(* IEC 61131-3 sources: REFUSR/GP/Refusr.jl/samples (part 13) *)

(* ---- 5-MUX_dozen-armor-usurp.st ---- *)
(*
This code implements a shuffled multiplexer with 5 control bits.
The control bits are: Data[N2], Data[N21], Data[N22], Data[N3], Data[N20]
The input bits are: Data[N24], Data[N4], Data[N27], Data[N1], Data[N23], Data[N25], Data[N5], Data[N26], Data[N31], Data[N7], Data[N8], Data[N6], Data[N9], Data[N28], Data[N13], Data[N11], Data[N12], Data[N29], Data[N30], Data[N33], Data[N10], Data[N34], Data[N35], Data[N37], Data[N32], Data[N14], Data[N16], Data[N36], Data[N17], Data[N18], Data[N19], Data[N15]

The symbolic expression is:
((((((((((((((((((((((((((((((((!(((((!(IN2)) & (!(IN21))) & (!(IN22))) & (!(IN3))) & (!(IN20)))) | IN24) & ((!((((IN2 & (!(IN21))) & (!(IN22))) & (!(IN3))) & (!(IN20)))) | IN4)) & ((!(((((!(IN2)) & IN21) & (!(IN22))) & (!(IN3))) & (!(IN20)))) | IN27)) & ((!((((IN2 & IN21) & (!(IN22))) & (!(IN3))) & (!(IN20)))) | IN1)) & ((!(((((!(IN2)) & (!(IN21))) & IN22) & (!(IN3))) & (!(IN20)))) | IN23)) & ((!((((IN2 & (!(IN21))) & IN22) & (!(IN3))) & (!(IN20)))) | IN25)) & ((!(((((!(IN2)) & IN21) & IN22) & (!(IN3))) & (!(IN20)))) | IN5)) & ((!((((IN2 & IN21) & IN22) & (!(IN3))) & (!(IN20)))) | IN26)) & ((!(((((!(IN2)) & (!(IN21))) & (!(IN22))) & IN3) & (!(IN20)))) | IN31)) & ((!((((IN2 & (!(IN21))) & (!(IN22))) & IN3) & (!(IN20)))) | IN7)) & ((!(((((!(IN2)) & IN21) & (!(IN22))) & IN3) & (!(IN20)))) | IN8)) & ((!((((IN2 & IN21) & (!(IN22))) & IN3) & (!(IN20)))) | IN6)) & ((!(((((!(IN2)) & (!(IN21))) & IN22) & IN3) & (!(IN20)))) | IN9)) & ((!((((IN2 & (!(IN21))) & IN22) & IN3) & (!(IN20)))) | IN28)) & ((!(((((!(IN2)) & IN21) & IN22) & IN3) & (!(IN20)))) | IN13)) & ((!((((IN2 & IN21) & IN22) & IN3) & (!(IN20)))) | IN11)) & ((!(((((!(IN2)) & (!(IN21))) & (!(IN22))) & (!(IN3))) & IN20)) | IN12)) & ((!((((IN2 & (!(IN21))) & (!(IN22))) & (!(IN3))) & IN20)) | IN29)) & ((!(((((!(IN2)) & IN21) & (!(IN22))) & (!(IN3))) & IN20)) | IN30)) & ((!((((IN2 & IN21) & (!(IN22))) & (!(IN3))) & IN20)) | IN33)) & ((!(((((!(IN2)) & (!(IN21))) & IN22) & (!(IN3))) & IN20)) | IN10)) & ((!((((IN2 & (!(IN21))) & IN22) & (!(IN3))) & IN20)) | IN34)) & ((!(((((!(IN2)) & IN21) & IN22) & (!(IN3))) & IN20)) | IN35)) & ((!((((IN2 & IN21) & IN22) & (!(IN3))) & IN20)) | IN37)) & ((!(((((!(IN2)) & (!(IN21))) & (!(IN22))) & IN3) & IN20)) | IN32)) & ((!((((IN2 & (!(IN21))) & (!(IN22))) & IN3) & IN20)) | IN14)) & ((!(((((!(IN2)) & IN21) & (!(IN22))) & IN3) & IN20)) | IN16)) & ((!((((IN2 & IN21) & (!(IN22))) & IN3) & IN20)) | IN36)) & ((!(((((!(IN2)) & (!(IN21))) & IN22) & IN3) & IN20)) | IN17)) & ((!((((IN2 & (!(IN21))) & IN22) & IN3) & IN20)) | IN18)) & ((!(((((!(IN2)) & IN21) & IN22) & IN3) & IN20)) | IN19)) & ((!((((IN2 & IN21) & IN22) & IN3) & IN20)) | IN15)

*)

FUNCTION_BLOCK F_CollectInput
  VAR_IN_OUT
      Data : ARRAY[1..40] OF BOOL;
  END_VAR
  VAR_INPUT
      TICK  : BOOL := 0;
      IN1   : BOOL := 0;
      IN2   : BOOL := 0;
      IN3   : BOOL := 0;
      IN4   : BOOL := 0;
      IN5   : BOOL := 0;
      RESET : BOOL := FALSE;
  END_VAR
  VAR_OUTPUT
      Finished : BOOL;
  END_VAR
  VAR
      j    : USINT := 1;
      tock : BOOL  := 0;
  END_VAR
  IF NOT RESET AND tock = NOT TICK THEN
      Data[j]   := IN1;
      Data[j+1] := IN2;
      Data[j+2] := IN3;
      Data[j+3] := IN4;
      Data[j+4] := IN5;
      j := j + 5;
      tock := TICK;
  ELSE
      j := 1;
      tock := 0;
  END_IF;
  Finished := (j > 40);
END_FUNCTION_BLOCK

PROGRAM Boiler
  VAR
    Data  : ARRAY[1..40] OF BOOL;
    Ready : BOOL;
    CollectInput : F_CollectInput;
  END_VAR
  VAR
    TICK     AT %IX1.0 : BOOL;
    IN1      AT %IX0.3 : BOOL;
    IN2      AT %IX0.4 : BOOL;
    IN3      AT %IX0.5 : BOOL;
    IN4      AT %IX0.6 : BOOL;
    IN5      AT %IX0.7 : BOOL;
    OutReady AT %QX0.0 : BOOL := FALSE;
    FeedNext AT %QX0.1 : BOOL := FALSE;
    Out      AT %QX0.2 : BOOL;
  END_VAR
  CollectInput(TICK:=TICK, IN1:=IN1, IN2:=IN2, IN3:=IN3, IN4:=IN4, IN5:=IN5);
  Ready := CollectInput.Finished;
  FeedNext := 1;
  IF Ready THEN
    Out := (((((((((((((((((((((((((((((((((NOT (((((NOT Data[2]) AND (NOT Data[21])) AND (NOT Data[22])) AND (NOT Data[3])) AND (NOT Data[20]))) OR Data[24]) AND ((NOT ((((Data[2] AND (NOT Data[21])) AND (NOT Data[22])) AND (NOT Data[3])) AND (NOT Data[20]))) OR Data[4])) AND ((NOT (((((NOT Data[2]) AND Data[21]) AND (NOT Data[22])) AND (NOT Data[3])) AND (NOT Data[20]))) OR Data[27])) AND ((NOT ((((Data[2] AND Data[21]) AND (NOT Data[22])) AND (NOT Data[3])) AND (NOT Data[20]))) OR Data[1])) AND ((NOT (((((NOT Data[2]) AND (NOT Data[21])) AND Data[22]) AND (NOT Data[3])) AND (NOT Data[20]))) OR Data[23])) AND ((NOT ((((Data[2] AND (NOT Data[21])) AND Data[22]) AND (NOT Data[3])) AND (NOT Data[20]))) OR Data[25])) AND ((NOT (((((NOT Data[2]) AND Data[21]) AND Data[22]) AND (NOT Data[3])) AND (NOT Data[20]))) OR Data[5])) AND ((NOT ((((Data[2] AND Data[21]) AND Data[22]) AND (NOT Data[3])) AND (NOT Data[20]))) OR Data[26])) AND ((NOT (((((NOT Data[2]) AND (NOT Data[21])) AND (NOT Data[22])) AND Data[3]) AND (NOT Data[20]))) OR Data[31])) AND ((NOT ((((Data[2] AND (NOT Data[21])) AND (NOT Data[22])) AND Data[3]) AND (NOT Data[20]))) OR Data[7])) AND ((NOT (((((NOT Data[2]) AND Data[21]) AND (NOT Data[22])) AND Data[3]) AND (NOT Data[20]))) OR Data[8])) AND ((NOT ((((Data[2] AND Data[21]) AND (NOT Data[22])) AND Data[3]) AND (NOT Data[20]))) OR Data[6])) AND ((NOT (((((NOT Data[2]) AND (NOT Data[21])) AND Data[22]) AND Data[3]) AND (NOT Data[20]))) OR Data[9])) AND ((NOT ((((Data[2] AND (NOT Data[21])) AND Data[22]) AND Data[3]) AND (NOT Data[20]))) OR Data[28])) AND ((NOT (((((NOT Data[2]) AND Data[21]) AND Data[22]) AND Data[3]) AND (NOT Data[20]))) OR Data[13])) AND ((NOT ((((Data[2] AND Data[21]) AND Data[22]) AND Data[3]) AND (NOT Data[20]))) OR Data[11])) AND ((NOT (((((NOT Data[2]) AND (NOT Data[21])) AND (NOT Data[22])) AND (NOT Data[3])) AND Data[20])) OR Data[12])) AND ((NOT ((((Data[2] AND (NOT Data[21])) AND (NOT Data[22])) AND (NOT Data[3])) AND Data[20])) OR Data[29])) AND ((NOT (((((NOT Data[2]) AND Data[21]) AND (NOT Data[22])) AND (NOT Data[3])) AND Data[20])) OR Data[30])) AND ((NOT ((((Data[2] AND Data[21]) AND (NOT Data[22])) AND (NOT Data[3])) AND Data[20])) OR Data[33])) AND ((NOT (((((NOT Data[2]) AND (NOT Data[21])) AND Data[22]) AND (NOT Data[3])) AND Data[20])) OR Data[10])) AND ((NOT ((((Data[2] AND (NOT Data[21])) AND Data[22]) AND (NOT Data[3])) AND Data[20])) OR Data[34])) AND ((NOT (((((NOT Data[2]) AND Data[21]) AND Data[22]) AND (NOT Data[3])) AND Data[20])) OR Data[35])) AND ((NOT ((((Data[2] AND Data[21]) AND Data[22]) AND (NOT Data[3])) AND Data[20])) OR Data[37])) AND ((NOT (((((NOT Data[2]) AND (NOT Data[21])) AND (NOT Data[22])) AND Data[3]) AND Data[20])) OR Data[32])) AND ((NOT ((((Data[2] AND (NOT Data[21])) AND (NOT Data[22])) AND Data[3]) AND Data[20])) OR Data[14])) AND ((NOT (((((NOT Data[2]) AND Data[21]) AND (NOT Data[22])) AND Data[3]) AND Data[20])) OR Data[16])) AND ((NOT ((((Data[2] AND Data[21]) AND (NOT Data[22])) AND Data[3]) AND Data[20])) OR Data[36])) AND ((NOT (((((NOT Data[2]) AND (NOT Data[21])) AND Data[22]) AND Data[3]) AND Data[20])) OR Data[17])) AND ((NOT ((((Data[2] AND (NOT Data[21])) AND Data[22]) AND Data[3]) AND Data[20])) OR Data[18])) AND ((NOT (((((NOT Data[2]) AND Data[21]) AND Data[22]) AND Data[3]) AND Data[20])) OR Data[19])) AND ((NOT ((((Data[2] AND Data[21]) AND Data[22]) AND Data[3]) AND Data[20])) OR Data[15]));
    OutReady := 1;
    CollectInput(RESET:=TRUE);
  END_IF;
END_PROGRAM

CONFIGURATION Config0
  RESOURCE Res0 ON PLC
    TASK task0(INTERVAL := T#20ms,PRIORITY := 0);
    PROGRAM instance0 WITH task0 : Boiler;
  END_RESOURCE
END_CONFIGURATION

(* ---- 5-MUX_froth-crick-hertz.st ---- *)
(*
This code implements a shuffled multiplexer with 5 control bits.
The control bits are: Data[N3], Data[N1], Data[N5], Data[N21], Data[N6]
The input bits are: Data[N4], Data[N20], Data[N2], Data[N7], Data[N22], Data[N8], Data[N10], Data[N11], Data[N13], Data[N26], Data[N23], Data[N25], Data[N9], Data[N14], Data[N24], Data[N29], Data[N16], Data[N27], Data[N15], Data[N12], Data[N17], Data[N19], Data[N32], Data[N30], Data[N28], Data[N18], Data[N31], Data[N33], Data[N37], Data[N35], Data[N36], Data[N34]

The symbolic expression is:
((((((((((((((((((((((((((((((((!(((((!(IN3)) & (!(IN1))) & (!(IN5))) & (!(IN21))) & (!(IN6)))) | IN4) & ((!((((IN3 & (!(IN1))) & (!(IN5))) & (!(IN21))) & (!(IN6)))) | IN20)) & ((!(((((!(IN3)) & IN1) & (!(IN5))) & (!(IN21))) & (!(IN6)))) | IN2)) & ((!((((IN3 & IN1) & (!(IN5))) & (!(IN21))) & (!(IN6)))) | IN7)) & ((!(((((!(IN3)) & (!(IN1))) & IN5) & (!(IN21))) & (!(IN6)))) | IN22)) & ((!((((IN3 & (!(IN1))) & IN5) & (!(IN21))) & (!(IN6)))) | IN8)) & ((!(((((!(IN3)) & IN1) & IN5) & (!(IN21))) & (!(IN6)))) | IN10)) & ((!((((IN3 & IN1) & IN5) & (!(IN21))) & (!(IN6)))) | IN11)) & ((!(((((!(IN3)) & (!(IN1))) & (!(IN5))) & IN21) & (!(IN6)))) | IN13)) & ((!((((IN3 & (!(IN1))) & (!(IN5))) & IN21) & (!(IN6)))) | IN26)) & ((!(((((!(IN3)) & IN1) & (!(IN5))) & IN21) & (!(IN6)))) | IN23)) & ((!((((IN3 & IN1) & (!(IN5))) & IN21) & (!(IN6)))) | IN25)) & ((!(((((!(IN3)) & (!(IN1))) & IN5) & IN21) & (!(IN6)))) | IN9)) & ((!((((IN3 & (!(IN1))) & IN5) & IN21) & (!(IN6)))) | IN14)) & ((!(((((!(IN3)) & IN1) & IN5) & IN21) & (!(IN6)))) | IN24)) & ((!((((IN3 & IN1) & IN5) & IN21) & (!(IN6)))) | IN29)) & ((!(((((!(IN3)) & (!(IN1))) & (!(IN5))) & (!(IN21))) & IN6)) | IN16)) & ((!((((IN3 & (!(IN1))) & (!(IN5))) & (!(IN21))) & IN6)) | IN27)) & ((!(((((!(IN3)) & IN1) & (!(IN5))) & (!(IN21))) & IN6)) | IN15)) & ((!((((IN3 & IN1) & (!(IN5))) & (!(IN21))) & IN6)) | IN12)) & ((!(((((!(IN3)) & (!(IN1))) & IN5) & (!(IN21))) & IN6)) | IN17)) & ((!((((IN3 & (!(IN1))) & IN5) & (!(IN21))) & IN6)) | IN19)) & ((!(((((!(IN3)) & IN1) & IN5) & (!(IN21))) & IN6)) | IN32)) & ((!((((IN3 & IN1) & IN5) & (!(IN21))) & IN6)) | IN30)) & ((!(((((!(IN3)) & (!(IN1))) & (!(IN5))) & IN21) & IN6)) | IN28)) & ((!((((IN3 & (!(IN1))) & (!(IN5))) & IN21) & IN6)) | IN18)) & ((!(((((!(IN3)) & IN1) & (!(IN5))) & IN21) & IN6)) | IN31)) & ((!((((IN3 & IN1) & (!(IN5))) & IN21) & IN6)) | IN33)) & ((!(((((!(IN3)) & (!(IN1))) & IN5) & IN21) & IN6)) | IN37)) & ((!((((IN3 & (!(IN1))) & IN5) & IN21) & IN6)) | IN35)) & ((!(((((!(IN3)) & IN1) & IN5) & IN21) & IN6)) | IN36)) & ((!((((IN3 & IN1) & IN5) & IN21) & IN6)) | IN34)

*)

FUNCTION_BLOCK F_CollectInput
  VAR_IN_OUT
      Data : ARRAY[1..40] OF BOOL;
  END_VAR
  VAR_INPUT
      TICK  : BOOL := 0;
      IN1   : BOOL := 0;
      IN2   : BOOL := 0;
      IN3   : BOOL := 0;
      IN4   : BOOL := 0;
      IN5   : BOOL := 0;
      RESET : BOOL := FALSE;
  END_VAR
  VAR_OUTPUT
      Finished : BOOL;
  END_VAR
  VAR
      j    : USINT := 1;
      tock : BOOL  := 0;
  END_VAR
  IF NOT RESET AND tock = NOT TICK THEN
      Data[j]   := IN1;
      Data[j+1] := IN2;
      Data[j+2] := IN3;
      Data[j+3] := IN4;
      Data[j+4] := IN5;
      j := j + 5;
      tock := TICK;
  ELSE
      j := 1;
      tock := 0;
  END_IF;
  Finished := (j > 40);
END_FUNCTION_BLOCK

PROGRAM Boiler
  VAR
    Data  : ARRAY[1..40] OF BOOL;
    Ready : BOOL;
    CollectInput : F_CollectInput;
  END_VAR
  VAR
    TICK     AT %IX1.0 : BOOL;
    IN1      AT %IX0.3 : BOOL;
    IN2      AT %IX0.4 : BOOL;
    IN3      AT %IX0.5 : BOOL;
    IN4      AT %IX0.6 : BOOL;
    IN5      AT %IX0.7 : BOOL;
    OutReady AT %QX0.0 : BOOL := FALSE;
    FeedNext AT %QX0.1 : BOOL := FALSE;
    Out      AT %QX0.2 : BOOL;
  END_VAR
  CollectInput(TICK:=TICK, IN1:=IN1, IN2:=IN2, IN3:=IN3, IN4:=IN4, IN5:=IN5);
  Ready := CollectInput.Finished;
  FeedNext := 1;
  IF Ready THEN
    Out := (((((((((((((((((((((((((((((((((NOT (((((NOT Data[3]) AND (NOT Data[1])) AND (NOT Data[5])) AND (NOT Data[21])) AND (NOT Data[6]))) OR Data[4]) AND ((NOT ((((Data[3] AND (NOT Data[1])) AND (NOT Data[5])) AND (NOT Data[21])) AND (NOT Data[6]))) OR Data[20])) AND ((NOT (((((NOT Data[3]) AND Data[1]) AND (NOT Data[5])) AND (NOT Data[21])) AND (NOT Data[6]))) OR Data[2])) AND ((NOT ((((Data[3] AND Data[1]) AND (NOT Data[5])) AND (NOT Data[21])) AND (NOT Data[6]))) OR Data[7])) AND ((NOT (((((NOT Data[3]) AND (NOT Data[1])) AND Data[5]) AND (NOT Data[21])) AND (NOT Data[6]))) OR Data[22])) AND ((NOT ((((Data[3] AND (NOT Data[1])) AND Data[5]) AND (NOT Data[21])) AND (NOT Data[6]))) OR Data[8])) AND ((NOT (((((NOT Data[3]) AND Data[1]) AND Data[5]) AND (NOT Data[21])) AND (NOT Data[6]))) OR Data[10])) AND ((NOT ((((Data[3] AND Data[1]) AND Data[5]) AND (NOT Data[21])) AND (NOT Data[6]))) OR Data[11])) AND ((NOT (((((NOT Data[3]) AND (NOT Data[1])) AND (NOT Data[5])) AND Data[21]) AND (NOT Data[6]))) OR Data[13])) AND ((NOT ((((Data[3] AND (NOT Data[1])) AND (NOT Data[5])) AND Data[21]) AND (NOT Data[6]))) OR Data[26])) AND ((NOT (((((NOT Data[3]) AND Data[1]) AND (NOT Data[5])) AND Data[21]) AND (NOT Data[6]))) OR Data[23])) AND ((NOT ((((Data[3] AND Data[1]) AND (NOT Data[5])) AND Data[21]) AND (NOT Data[6]))) OR Data[25])) AND ((NOT (((((NOT Data[3]) AND (NOT Data[1])) AND Data[5]) AND Data[21]) AND (NOT Data[6]))) OR Data[9])) AND ((NOT ((((Data[3] AND (NOT Data[1])) AND Data[5]) AND Data[21]) AND (NOT Data[6]))) OR Data[14])) AND ((NOT (((((NOT Data[3]) AND Data[1]) AND Data[5]) AND Data[21]) AND (NOT Data[6]))) OR Data[24])) AND ((NOT ((((Data[3] AND Data[1]) AND Data[5]) AND Data[21]) AND (NOT Data[6]))) OR Data[29])) AND ((NOT (((((NOT Data[3]) AND (NOT Data[1])) AND (NOT Data[5])) AND (NOT Data[21])) AND Data[6])) OR Data[16])) AND ((NOT ((((Data[3] AND (NOT Data[1])) AND (NOT Data[5])) AND (NOT Data[21])) AND Data[6])) OR Data[27])) AND ((NOT (((((NOT Data[3]) AND Data[1]) AND (NOT Data[5])) AND (NOT Data[21])) AND Data[6])) OR Data[15])) AND ((NOT ((((Data[3] AND Data[1]) AND (NOT Data[5])) AND (NOT Data[21])) AND Data[6])) OR Data[12])) AND ((NOT (((((NOT Data[3]) AND (NOT Data[1])) AND Data[5]) AND (NOT Data[21])) AND Data[6])) OR Data[17])) AND ((NOT ((((Data[3] AND (NOT Data[1])) AND Data[5]) AND (NOT Data[21])) AND Data[6])) OR Data[19])) AND ((NOT (((((NOT Data[3]) AND Data[1]) AND Data[5]) AND (NOT Data[21])) AND Data[6])) OR Data[32])) AND ((NOT ((((Data[3] AND Data[1]) AND Data[5]) AND (NOT Data[21])) AND Data[6])) OR Data[30])) AND ((NOT (((((NOT Data[3]) AND (NOT Data[1])) AND (NOT Data[5])) AND Data[21]) AND Data[6])) OR Data[28])) AND ((NOT ((((Data[3] AND (NOT Data[1])) AND (NOT Data[5])) AND Data[21]) AND Data[6])) OR Data[18])) AND ((NOT (((((NOT Data[3]) AND Data[1]) AND (NOT Data[5])) AND Data[21]) AND Data[6])) OR Data[31])) AND ((NOT ((((Data[3] AND Data[1]) AND (NOT Data[5])) AND Data[21]) AND Data[6])) OR Data[33])) AND ((NOT (((((NOT Data[3]) AND (NOT Data[1])) AND Data[5]) AND Data[21]) AND Data[6])) OR Data[37])) AND ((NOT ((((Data[3] AND (NOT Data[1])) AND Data[5]) AND Data[21]) AND Data[6])) OR Data[35])) AND ((NOT (((((NOT Data[3]) AND Data[1]) AND Data[5]) AND Data[21]) AND Data[6])) OR Data[36])) AND ((NOT ((((Data[3] AND Data[1]) AND Data[5]) AND Data[21]) AND Data[6])) OR Data[34]));
    OutReady := 1;
    CollectInput(RESET:=TRUE);
  END_IF;
END_PROGRAM

CONFIGURATION Config0
  RESOURCE Res0 ON PLC
    TASK task0(INTERVAL := T#20ms,PRIORITY := 0);
    PROGRAM instance0 WITH task0 : Boiler;
  END_RESOURCE
END_CONFIGURATION

(* ---- 5-MUX_funds-axman-titan.st ---- *)
(*
This code implements a shuffled multiplexer with 5 control bits.
The control bits are: Data[N22], Data[N1], Data[N23], Data[N20], Data[N24]
The input bits are: Data[N26], Data[N21], Data[N29], Data[N27], Data[N7], Data[N4], Data[N30], Data[N33], Data[N25], Data[N28], Data[N31], Data[N34], Data[N6], Data[N2], Data[N32], Data[N8], Data[N3], Data[N14], Data[N9], Data[N5], Data[N10], Data[N35], Data[N12], Data[N13], Data[N16], Data[N15], Data[N36], Data[N37], Data[N11], Data[N17], Data[N19], Data[N18]

The symbolic expression is:
((((((((((((((((((((((((((((((((!(((((!(IN22)) & (!(IN1))) & (!(IN23))) & (!(IN20))) & (!(IN24)))) | IN26) & ((!((((IN22 & (!(IN1))) & (!(IN23))) & (!(IN20))) & (!(IN24)))) | IN21)) & ((!(((((!(IN22)) & IN1) & (!(IN23))) & (!(IN20))) & (!(IN24)))) | IN29)) & ((!((((IN22 & IN1) & (!(IN23))) & (!(IN20))) & (!(IN24)))) | IN27)) & ((!(((((!(IN22)) & (!(IN1))) & IN23) & (!(IN20))) & (!(IN24)))) | IN7)) & ((!((((IN22 & (!(IN1))) & IN23) & (!(IN20))) & (!(IN24)))) | IN4)) & ((!(((((!(IN22)) & IN1) & IN23) & (!(IN20))) & (!(IN24)))) | IN30)) & ((!((((IN22 & IN1) & IN23) & (!(IN20))) & (!(IN24)))) | IN33)) & ((!(((((!(IN22)) & (!(IN1))) & (!(IN23))) & IN20) & (!(IN24)))) | IN25)) & ((!((((IN22 & (!(IN1))) & (!(IN23))) & IN20) & (!(IN24)))) | IN28)) & ((!(((((!(IN22)) & IN1) & (!(IN23))) & IN20) & (!(IN24)))) | IN31)) & ((!((((IN22 & IN1) & (!(IN23))) & IN20) & (!(IN24)))) | IN34)) & ((!(((((!(IN22)) & (!(IN1))) & IN23) & IN20) & (!(IN24)))) | IN6)) & ((!((((IN22 & (!(IN1))) & IN23) & IN20) & (!(IN24)))) | IN2)) & ((!(((((!(IN22)) & IN1) & IN23) & IN20) & (!(IN24)))) | IN32)) & ((!((((IN22 & IN1) & IN23) & IN20) & (!(IN24)))) | IN8)) & ((!(((((!(IN22)) & (!(IN1))) & (!(IN23))) & (!(IN20))) & IN24)) | IN3)) & ((!((((IN22 & (!(IN1))) & (!(IN23))) & (!(IN20))) & IN24)) | IN14)) & ((!(((((!(IN22)) & IN1) & (!(IN23))) & (!(IN20))) & IN24)) | IN9)) & ((!((((IN22 & IN1) & (!(IN23))) & (!(IN20))) & IN24)) | IN5)) & ((!(((((!(IN22)) & (!(IN1))) & IN23) & (!(IN20))) & IN24)) | IN10)) & ((!((((IN22 & (!(IN1))) & IN23) & (!(IN20))) & IN24)) | IN35)) & ((!(((((!(IN22)) & IN1) & IN23) & (!(IN20))) & IN24)) | IN12)) & ((!((((IN22 & IN1) & IN23) & (!(IN20))) & IN24)) | IN13)) & ((!(((((!(IN22)) & (!(IN1))) & (!(IN23))) & IN20) & IN24)) | IN16)) & ((!((((IN22 & (!(IN1))) & (!(IN23))) & IN20) & IN24)) | IN15)) & ((!(((((!(IN22)) & IN1) & (!(IN23))) & IN20) & IN24)) | IN36)) & ((!((((IN22 & IN1) & (!(IN23))) & IN20) & IN24)) | IN37)) & ((!(((((!(IN22)) & (!(IN1))) & IN23) & IN20) & IN24)) | IN11)) & ((!((((IN22 & (!(IN1))) & IN23) & IN20) & IN24)) | IN17)) & ((!(((((!(IN22)) & IN1) & IN23) & IN20) & IN24)) | IN19)) & ((!((((IN22 & IN1) & IN23) & IN20) & IN24)) | IN18)

*)

FUNCTION_BLOCK F_CollectInput
  VAR_IN_OUT
      Data : ARRAY[1..40] OF BOOL;
  END_VAR
  VAR_INPUT
      TICK  : BOOL := 0;
      IN1   : BOOL := 0;
      IN2   : BOOL := 0;
      IN3   : BOOL := 0;
      IN4   : BOOL := 0;
      IN5   : BOOL := 0;
      RESET : BOOL := FALSE;
  END_VAR
  VAR_OUTPUT
      Finished : BOOL;
  END_VAR
  VAR
      j    : USINT := 1;
      tock : BOOL  := 0;
  END_VAR
  IF NOT RESET AND tock = NOT TICK THEN
      Data[j]   := IN1;
      Data[j+1] := IN2;
      Data[j+2] := IN3;
      Data[j+3] := IN4;
      Data[j+4] := IN5;
      j := j + 5;
      tock := TICK;
  ELSE
      j := 1;
      tock := 0;
  END_IF;
  Finished := (j > 40);
END_FUNCTION_BLOCK

PROGRAM Boiler
  VAR
    Data  : ARRAY[1..40] OF BOOL;
    Ready : BOOL;
    CollectInput : F_CollectInput;
  END_VAR
  VAR
    TICK     AT %IX1.0 : BOOL;
    IN1      AT %IX0.3 : BOOL;
    IN2      AT %IX0.4 : BOOL;
    IN3      AT %IX0.5 : BOOL;
    IN4      AT %IX0.6 : BOOL;
    IN5      AT %IX0.7 : BOOL;
    OutReady AT %QX0.0 : BOOL := FALSE;
    FeedNext AT %QX0.1 : BOOL := FALSE;
    Out      AT %QX0.2 : BOOL;
  END_VAR
  CollectInput(TICK:=TICK, IN1:=IN1, IN2:=IN2, IN3:=IN3, IN4:=IN4, IN5:=IN5);
  Ready := CollectInput.Finished;
  FeedNext := 1;
  IF Ready THEN
    Out := (((((((((((((((((((((((((((((((((NOT (((((NOT Data[22]) AND (NOT Data[1])) AND (NOT Data[23])) AND (NOT Data[20])) AND (NOT Data[24]))) OR Data[26]) AND ((NOT ((((Data[22] AND (NOT Data[1])) AND (NOT Data[23])) AND (NOT Data[20])) AND (NOT Data[24]))) OR Data[21])) AND ((NOT (((((NOT Data[22]) AND Data[1]) AND (NOT Data[23])) AND (NOT Data[20])) AND (NOT Data[24]))) OR Data[29])) AND ((NOT ((((Data[22] AND Data[1]) AND (NOT Data[23])) AND (NOT Data[20])) AND (NOT Data[24]))) OR Data[27])) AND ((NOT (((((NOT Data[22]) AND (NOT Data[1])) AND Data[23]) AND (NOT Data[20])) AND (NOT Data[24]))) OR Data[7])) AND ((NOT ((((Data[22] AND (NOT Data[1])) AND Data[23]) AND (NOT Data[20])) AND (NOT Data[24]))) OR Data[4])) AND ((NOT (((((NOT Data[22]) AND Data[1]) AND Data[23]) AND (NOT Data[20])) AND (NOT Data[24]))) OR Data[30])) AND ((NOT ((((Data[22] AND Data[1]) AND Data[23]) AND (NOT Data[20])) AND (NOT Data[24]))) OR Data[33])) AND ((NOT (((((NOT Data[22]) AND (NOT Data[1])) AND (NOT Data[23])) AND Data[20]) AND (NOT Data[24]))) OR Data[25])) AND ((NOT ((((Data[22] AND (NOT Data[1])) AND (NOT Data[23])) AND Data[20]) AND (NOT Data[24]))) OR Data[28])) AND ((NOT (((((NOT Data[22]) AND Data[1]) AND (NOT Data[23])) AND Data[20]) AND (NOT Data[24]))) OR Data[31])) AND ((NOT ((((Data[22] AND Data[1]) AND (NOT Data[23])) AND Data[20]) AND (NOT Data[24]))) OR Data[34])) AND ((NOT (((((NOT Data[22]) AND (NOT Data[1])) AND Data[23]) AND Data[20]) AND (NOT Data[24]))) OR Data[6])) AND ((NOT ((((Data[22] AND (NOT Data[1])) AND Data[23]) AND Data[20]) AND (NOT Data[24]))) OR Data[2])) AND ((NOT (((((NOT Data[22]) AND Data[1]) AND Data[23]) AND Data[20]) AND (NOT Data[24]))) OR Data[32])) AND ((NOT ((((Data[22] AND Data[1]) AND Data[23]) AND Data[20]) AND (NOT Data[24]))) OR Data[8])) AND ((NOT (((((NOT Data[22]) AND (NOT Data[1])) AND (NOT Data[23])) AND (NOT Data[20])) AND Data[24])) OR Data[3])) AND ((NOT ((((Data[22] AND (NOT Data[1])) AND (NOT Data[23])) AND (NOT Data[20])) AND Data[24])) OR Data[14])) AND ((NOT (((((NOT Data[22]) AND Data[1]) AND (NOT Data[23])) AND (NOT Data[20])) AND Data[24])) OR Data[9])) AND ((NOT ((((Data[22] AND Data[1]) AND (NOT Data[23])) AND (NOT Data[20])) AND Data[24])) OR Data[5])) AND ((NOT (((((NOT Data[22]) AND (NOT Data[1])) AND Data[23]) AND (NOT Data[20])) AND Data[24])) OR Data[10])) AND ((NOT ((((Data[22] AND (NOT Data[1])) AND Data[23]) AND (NOT Data[20])) AND Data[24])) OR Data[35])) AND ((NOT (((((NOT Data[22]) AND Data[1]) AND Data[23]) AND (NOT Data[20])) AND Data[24])) OR Data[12])) AND ((NOT ((((Data[22] AND Data[1]) AND Data[23]) AND (NOT Data[20])) AND Data[24])) OR Data[13])) AND ((NOT (((((NOT Data[22]) AND (NOT Data[1])) AND (NOT Data[23])) AND Data[20]) AND Data[24])) OR Data[16])) AND ((NOT ((((Data[22] AND (NOT Data[1])) AND (NOT Data[23])) AND Data[20]) AND Data[24])) OR Data[15])) AND ((NOT (((((NOT Data[22]) AND Data[1]) AND (NOT Data[23])) AND Data[20]) AND Data[24])) OR Data[36])) AND ((NOT ((((Data[22] AND Data[1]) AND (NOT Data[23])) AND Data[20]) AND Data[24])) OR Data[37])) AND ((NOT (((((NOT Data[22]) AND (NOT Data[1])) AND Data[23]) AND Data[20]) AND Data[24])) OR Data[11])) AND ((NOT ((((Data[22] AND (NOT Data[1])) AND Data[23]) AND Data[20]) AND Data[24])) OR Data[17])) AND ((NOT (((((NOT Data[22]) AND Data[1]) AND Data[23]) AND Data[20]) AND Data[24])) OR Data[19])) AND ((NOT ((((Data[22] AND Data[1]) AND Data[23]) AND Data[20]) AND Data[24])) OR Data[18]));
    OutReady := 1;
    CollectInput(RESET:=TRUE);
  END_IF;
END_PROGRAM

CONFIGURATION Config0
  RESOURCE Res0 ON PLC
    TASK task0(INTERVAL := T#20ms,PRIORITY := 0);
    PROGRAM instance0 WITH task0 : Boiler;
  END_RESOURCE
END_CONFIGURATION

(* ---- 5-MUX_fungi-exalt-steer.st ---- *)
(*
This code implements a shuffled multiplexer with 5 control bits.
The control bits are: Data[N1], Data[N3], Data[N5], Data[N2], Data[N21]
The input bits are: Data[N20], Data[N25], Data[N6], Data[N23], Data[N26], Data[N24], Data[N4], Data[N13], Data[N28], Data[N7], Data[N22], Data[N29], Data[N30], Data[N27], Data[N10], Data[N11], Data[N31], Data[N33], Data[N34], Data[N32], Data[N8], Data[N36], Data[N35], Data[N37], Data[N15], Data[N17], Data[N14], Data[N9], Data[N12], Data[N18], Data[N16], Data[N19]

The symbolic expression is:
((((((((((((((((((((((((((((((((!(((((!(IN1)) & (!(IN3))) & (!(IN5))) & (!(IN2))) & (!(IN21)))) | IN20) & ((!((((IN1 & (!(IN3))) & (!(IN5))) & (!(IN2))) & (!(IN21)))) | IN25)) & ((!(((((!(IN1)) & IN3) & (!(IN5))) & (!(IN2))) & (!(IN21)))) | IN6)) & ((!((((IN1 & IN3) & (!(IN5))) & (!(IN2))) & (!(IN21)))) | IN23)) & ((!(((((!(IN1)) & (!(IN3))) & IN5) & (!(IN2))) & (!(IN21)))) | IN26)) & ((!((((IN1 & (!(IN3))) & IN5) & (!(IN2))) & (!(IN21)))) | IN24)) & ((!(((((!(IN1)) & IN3) & IN5) & (!(IN2))) & (!(IN21)))) | IN4)) & ((!((((IN1 & IN3) & IN5) & (!(IN2))) & (!(IN21)))) | IN13)) & ((!(((((!(IN1)) & (!(IN3))) & (!(IN5))) & IN2) & (!(IN21)))) | IN28)) & ((!((((IN1 & (!(IN3))) & (!(IN5))) & IN2) & (!(IN21)))) | IN7)) & ((!(((((!(IN1)) & IN3) & (!(IN5))) & IN2) & (!(IN21)))) | IN22)) & ((!((((IN1 & IN3) & (!(IN5))) & IN2) & (!(IN21)))) | IN29)) & ((!(((((!(IN1)) & (!(IN3))) & IN5) & IN2) & (!(IN21)))) | IN30)) & ((!((((IN1 & (!(IN3))) & IN5) & IN2) & (!(IN21)))) | IN27)) & ((!(((((!(IN1)) & IN3) & IN5) & IN2) & (!(IN21)))) | IN10)) & ((!((((IN1 & IN3) & IN5) & IN2) & (!(IN21)))) | IN11)) & ((!(((((!(IN1)) & (!(IN3))) & (!(IN5))) & (!(IN2))) & IN21)) | IN31)) & ((!((((IN1 & (!(IN3))) & (!(IN5))) & (!(IN2))) & IN21)) | IN33)) & ((!(((((!(IN1)) & IN3) & (!(IN5))) & (!(IN2))) & IN21)) | IN34)) & ((!((((IN1 & IN3) & (!(IN5))) & (!(IN2))) & IN21)) | IN32)) & ((!(((((!(IN1)) & (!(IN3))) & IN5) & (!(IN2))) & IN21)) | IN8)) & ((!((((IN1 & (!(IN3))) & IN5) & (!(IN2))) & IN21)) | IN36)) & ((!(((((!(IN1)) & IN3) & IN5) & (!(IN2))) & IN21)) | IN35)) & ((!((((IN1 & IN3) & IN5) & (!(IN2))) & IN21)) | IN37)) & ((!(((((!(IN1)) & (!(IN3))) & (!(IN5))) & IN2) & IN21)) | IN15)) & ((!((((IN1 & (!(IN3))) & (!(IN5))) & IN2) & IN21)) | IN17)) & ((!(((((!(IN1)) & IN3) & (!(IN5))) & IN2) & IN21)) | IN14)) & ((!((((IN1 & IN3) & (!(IN5))) & IN2) & IN21)) | IN9)) & ((!(((((!(IN1)) & (!(IN3))) & IN5) & IN2) & IN21)) | IN12)) & ((!((((IN1 & (!(IN3))) & IN5) & IN2) & IN21)) | IN18)) & ((!(((((!(IN1)) & IN3) & IN5) & IN2) & IN21)) | IN16)) & ((!((((IN1 & IN3) & IN5) & IN2) & IN21)) | IN19)

*)

FUNCTION_BLOCK F_CollectInput
  VAR_IN_OUT
      Data : ARRAY[1..40] OF BOOL;
  END_VAR
  VAR_INPUT
      TICK  : BOOL := 0;
      IN1   : BOOL := 0;
      IN2   : BOOL := 0;
      IN3   : BOOL := 0;
      IN4   : BOOL := 0;
      IN5   : BOOL := 0;
      RESET : BOOL := FALSE;
  END_VAR
  VAR_OUTPUT
      Finished : BOOL;
  END_VAR
  VAR
      j    : USINT := 1;
      tock : BOOL  := 0;
  END_VAR
  IF NOT RESET AND tock = NOT TICK THEN
      Data[j]   := IN1;
      Data[j+1] := IN2;
      Data[j+2] := IN3;
      Data[j+3] := IN4;
      Data[j+4] := IN5;
      j := j + 5;
      tock := TICK;
  ELSE
      j := 1;
      tock := 0;
  END_IF;
  Finished := (j > 40);
END_FUNCTION_BLOCK

PROGRAM Boiler
  VAR
    Data  : ARRAY[1..40] OF BOOL;
    Ready : BOOL;
    CollectInput : F_CollectInput;
  END_VAR
  VAR
    TICK     AT %IX1.0 : BOOL;
    IN1      AT %IX0.3 : BOOL;
    IN2      AT %IX0.4 : BOOL;
    IN3      AT %IX0.5 : BOOL;
    IN4      AT %IX0.6 : BOOL;
    IN5      AT %IX0.7 : BOOL;
    OutReady AT %QX0.0 : BOOL := FALSE;
    FeedNext AT %QX0.1 : BOOL := FALSE;
    Out      AT %QX0.2 : BOOL;
  END_VAR
  CollectInput(TICK:=TICK, IN1:=IN1, IN2:=IN2, IN3:=IN3, IN4:=IN4, IN5:=IN5);
  Ready := CollectInput.Finished;
  FeedNext := 1;
  IF Ready THEN
    Out := (((((((((((((((((((((((((((((((((NOT (((((NOT Data[1]) AND (NOT Data[3])) AND (NOT Data[5])) AND (NOT Data[2])) AND (NOT Data[21]))) OR Data[20]) AND ((NOT ((((Data[1] AND (NOT Data[3])) AND (NOT Data[5])) AND (NOT Data[2])) AND (NOT Data[21]))) OR Data[25])) AND ((NOT (((((NOT Data[1]) AND Data[3]) AND (NOT Data[5])) AND (NOT Data[2])) AND (NOT Data[21]))) OR Data[6])) AND ((NOT ((((Data[1] AND Data[3]) AND (NOT Data[5])) AND (NOT Data[2])) AND (NOT Data[21]))) OR Data[23])) AND ((NOT (((((NOT Data[1]) AND (NOT Data[3])) AND Data[5]) AND (NOT Data[2])) AND (NOT Data[21]))) OR Data[26])) AND ((NOT ((((Data[1] AND (NOT Data[3])) AND Data[5]) AND (NOT Data[2])) AND (NOT Data[21]))) OR Data[24])) AND ((NOT (((((NOT Data[1]) AND Data[3]) AND Data[5]) AND (NOT Data[2])) AND (NOT Data[21]))) OR Data[4])) AND ((NOT ((((Data[1] AND Data[3]) AND Data[5]) AND (NOT Data[2])) AND (NOT Data[21]))) OR Data[13])) AND ((NOT (((((NOT Data[1]) AND (NOT Data[3])) AND (NOT Data[5])) AND Data[2]) AND (NOT Data[21]))) OR Data[28])) AND ((NOT ((((Data[1] AND (NOT Data[3])) AND (NOT Data[5])) AND Data[2]) AND (NOT Data[21]))) OR Data[7])) AND ((NOT (((((NOT Data[1]) AND Data[3]) AND (NOT Data[5])) AND Data[2]) AND (NOT Data[21]))) OR Data[22])) AND ((NOT ((((Data[1] AND Data[3]) AND (NOT Data[5])) AND Data[2]) AND (NOT Data[21]))) OR Data[29])) AND ((NOT (((((NOT Data[1]) AND (NOT Data[3])) AND Data[5]) AND Data[2]) AND (NOT Data[21]))) OR Data[30])) AND ((NOT ((((Data[1] AND (NOT Data[3])) AND Data[5]) AND Data[2]) AND (NOT Data[21]))) OR Data[27])) AND ((NOT (((((NOT Data[1]) AND Data[3]) AND Data[5]) AND Data[2]) AND (NOT Data[21]))) OR Data[10])) AND ((NOT ((((Data[1] AND Data[3]) AND Data[5]) AND Data[2]) AND (NOT Data[21]))) OR Data[11])) AND ((NOT (((((NOT Data[1]) AND (NOT Data[3])) AND (NOT Data[5])) AND (NOT Data[2])) AND Data[21])) OR Data[31])) AND ((NOT ((((Data[1] AND (NOT Data[3])) AND (NOT Data[5])) AND (NOT Data[2])) AND Data[21])) OR Data[33])) AND ((NOT (((((NOT Data[1]) AND Data[3]) AND (NOT Data[5])) AND (NOT Data[2])) AND Data[21])) OR Data[34])) AND ((NOT ((((Data[1] AND Data[3]) AND (NOT Data[5])) AND (NOT Data[2])) AND Data[21])) OR Data[32])) AND ((NOT (((((NOT Data[1]) AND (NOT Data[3])) AND Data[5]) AND (NOT Data[2])) AND Data[21])) OR Data[8])) AND ((NOT ((((Data[1] AND (NOT Data[3])) AND Data[5]) AND (NOT Data[2])) AND Data[21])) OR Data[36])) AND ((NOT (((((NOT Data[1]) AND Data[3]) AND Data[5]) AND (NOT Data[2])) AND Data[21])) OR Data[35])) AND ((NOT ((((Data[1] AND Data[3]) AND Data[5]) AND (NOT Data[2])) AND Data[21])) OR Data[37])) AND ((NOT (((((NOT Data[1]) AND (NOT Data[3])) AND (NOT Data[5])) AND Data[2]) AND Data[21])) OR Data[15])) AND ((NOT ((((Data[1] AND (NOT Data[3])) AND (NOT Data[5])) AND Data[2]) AND Data[21])) OR Data[17])) AND ((NOT (((((NOT Data[1]) AND Data[3]) AND (NOT Data[5])) AND Data[2]) AND Data[21])) OR Data[14])) AND ((NOT ((((Data[1] AND Data[3]) AND (NOT Data[5])) AND Data[2]) AND Data[21])) OR Data[9])) AND ((NOT (((((NOT Data[1]) AND (NOT Data[3])) AND Data[5]) AND Data[2]) AND Data[21])) OR Data[12])) AND ((NOT ((((Data[1] AND (NOT Data[3])) AND Data[5]) AND Data[2]) AND Data[21])) OR Data[18])) AND ((NOT (((((NOT Data[1]) AND Data[3]) AND Data[5]) AND Data[2]) AND Data[21])) OR Data[16])) AND ((NOT ((((Data[1] AND Data[3]) AND Data[5]) AND Data[2]) AND Data[21])) OR Data[19]));
    OutReady := 1;
    CollectInput(RESET:=TRUE);
  END_IF;
END_PROGRAM

CONFIGURATION Config0
  RESOURCE Res0 ON PLC
    TASK task0(INTERVAL := T#20ms,PRIORITY := 0);
    PROGRAM instance0 WITH task0 : Boiler;
  END_RESOURCE
END_CONFIGURATION

(* ---- 5-MUX_gipsy-agave-shock.st ---- *)
(*
This code implements a shuffled multiplexer with 5 control bits.
The control bits are: Data[N21], Data[N23], Data[N24], Data[N25], Data[N26]
The input bits are: Data[N4], Data[N5], Data[N1], Data[N6], Data[N27], Data[N20], Data[N30], Data[N31], Data[N22], Data[N33], Data[N9], Data[N32], Data[N28], Data[N34], Data[N37], Data[N2], Data[N29], Data[N36], Data[N3], Data[N7], Data[N35], Data[N8], Data[N13], Data[N12], Data[N11], Data[N19], Data[N18], Data[N15], Data[N10], Data[N14], Data[N16], Data[N17]

The symbolic expression is:
((((((((((((((((((((((((((((((((!(((((!(IN21)) & (!(IN23))) & (!(IN24))) & (!(IN25))) & (!(IN26)))) | IN4) & ((!((((IN21 & (!(IN23))) & (!(IN24))) & (!(IN25))) & (!(IN26)))) | IN5)) & ((!(((((!(IN21)) & IN23) & (!(IN24))) & (!(IN25))) & (!(IN26)))) | IN1)) & ((!((((IN21 & IN23) & (!(IN24))) & (!(IN25))) & (!(IN26)))) | IN6)) & ((!(((((!(IN21)) & (!(IN23))) & IN24) & (!(IN25))) & (!(IN26)))) | IN27)) & ((!((((IN21 & (!(IN23))) & IN24) & (!(IN25))) & (!(IN26)))) | IN20)) & ((!(((((!(IN21)) & IN23) & IN24) & (!(IN25))) & (!(IN26)))) | IN30)) & ((!((((IN21 & IN23) & IN24) & (!(IN25))) & (!(IN26)))) | IN31)) & ((!(((((!(IN21)) & (!(IN23))) & (!(IN24))) & IN25) & (!(IN26)))) | IN22)) & ((!((((IN21 & (!(IN23))) & (!(IN24))) & IN25) & (!(IN26)))) | IN33)) & ((!(((((!(IN21)) & IN23) & (!(IN24))) & IN25) & (!(IN26)))) | IN9)) & ((!((((IN21 & IN23) & (!(IN24))) & IN25) & (!(IN26)))) | IN32)) & ((!(((((!(IN21)) & (!(IN23))) & IN24) & IN25) & (!(IN26)))) | IN28)) & ((!((((IN21 & (!(IN23))) & IN24) & IN25) & (!(IN26)))) | IN34)) & ((!(((((!(IN21)) & IN23) & IN24) & IN25) & (!(IN26)))) | IN37)) & ((!((((IN21 & IN23) & IN24) & IN25) & (!(IN26)))) | IN2)) & ((!(((((!(IN21)) & (!(IN23))) & (!(IN24))) & (!(IN25))) & IN26)) | IN29)) & ((!((((IN21 & (!(IN23))) & (!(IN24))) & (!(IN25))) & IN26)) | IN36)) & ((!(((((!(IN21)) & IN23) & (!(IN24))) & (!(IN25))) & IN26)) | IN3)) & ((!((((IN21 & IN23) & (!(IN24))) & (!(IN25))) & IN26)) | IN7)) & ((!(((((!(IN21)) & (!(IN23))) & IN24) & (!(IN25))) & IN26)) | IN35)) & ((!((((IN21 & (!(IN23))) & IN24) & (!(IN25))) & IN26)) | IN8)) & ((!(((((!(IN21)) & IN23) & IN24) & (!(IN25))) & IN26)) | IN13)) & ((!((((IN21 & IN23) & IN24) & (!(IN25))) & IN26)) | IN12)) & ((!(((((!(IN21)) & (!(IN23))) & (!(IN24))) & IN25) & IN26)) | IN11)) & ((!((((IN21 & (!(IN23))) & (!(IN24))) & IN25) & IN26)) | IN19)) & ((!(((((!(IN21)) & IN23) & (!(IN24))) & IN25) & IN26)) | IN18)) & ((!((((IN21 & IN23) & (!(IN24))) & IN25) & IN26)) | IN15)) & ((!(((((!(IN21)) & (!(IN23))) & IN24) & IN25) & IN26)) | IN10)) & ((!((((IN21 & (!(IN23))) & IN24) & IN25) & IN26)) | IN14)) & ((!(((((!(IN21)) & IN23) & IN24) & IN25) & IN26)) | IN16)) & ((!((((IN21 & IN23) & IN24) & IN25) & IN26)) | IN17)

*)

FUNCTION_BLOCK F_CollectInput
  VAR_IN_OUT
      Data : ARRAY[1..40] OF BOOL;
  END_VAR
  VAR_INPUT
      TICK  : BOOL := 0;
      IN1   : BOOL := 0;
      IN2   : BOOL := 0;
      IN3   : BOOL := 0;
      IN4   : BOOL := 0;
      IN5   : BOOL := 0;
      RESET : BOOL := FALSE;
  END_VAR
  VAR_OUTPUT
      Finished : BOOL;
  END_VAR
  VAR
      j    : USINT := 1;
      tock : BOOL  := 0;
  END_VAR
  IF NOT RESET AND tock = NOT TICK THEN
      Data[j]   := IN1;
      Data[j+1] := IN2;
      Data[j+2] := IN3;
      Data[j+3] := IN4;
      Data[j+4] := IN5;
      j := j + 5;
      tock := TICK;
  ELSE
      j := 1;
      tock := 0;
  END_IF;
  Finished := (j > 40);
END_FUNCTION_BLOCK

PROGRAM Boiler
  VAR
    Data  : ARRAY[1..40] OF BOOL;
    Ready : BOOL;
    CollectInput : F_CollectInput;
  END_VAR
  VAR
    TICK     AT %IX1.0 : BOOL;
    IN1      AT %IX0.3 : BOOL;
    IN2      AT %IX0.4 : BOOL;
    IN3      AT %IX0.5 : BOOL;
    IN4      AT %IX0.6 : BOOL;
    IN5      AT %IX0.7 : BOOL;
    OutReady AT %QX0.0 : BOOL := FALSE;
    FeedNext AT %QX0.1 : BOOL := FALSE;
    Out      AT %QX0.2 : BOOL;
  END_VAR
  CollectInput(TICK:=TICK, IN1:=IN1, IN2:=IN2, IN3:=IN3, IN4:=IN4, IN5:=IN5);
  Ready := CollectInput.Finished;
  FeedNext := 1;
  IF Ready THEN
    Out := (((((((((((((((((((((((((((((((((NOT (((((NOT Data[21]) AND (NOT Data[23])) AND (NOT Data[24])) AND (NOT Data[25])) AND (NOT Data[26]))) OR Data[4]) AND ((NOT ((((Data[21] AND (NOT Data[23])) AND (NOT Data[24])) AND (NOT Data[25])) AND (NOT Data[26]))) OR Data[5])) AND ((NOT (((((NOT Data[21]) AND Data[23]) AND (NOT Data[24])) AND (NOT Data[25])) AND (NOT Data[26]))) OR Data[1])) AND ((NOT ((((Data[21] AND Data[23]) AND (NOT Data[24])) AND (NOT Data[25])) AND (NOT Data[26]))) OR Data[6])) AND ((NOT (((((NOT Data[21]) AND (NOT Data[23])) AND Data[24]) AND (NOT Data[25])) AND (NOT Data[26]))) OR Data[27])) AND ((NOT ((((Data[21] AND (NOT Data[23])) AND Data[24]) AND (NOT Data[25])) AND (NOT Data[26]))) OR Data[20])) AND ((NOT (((((NOT Data[21]) AND Data[23]) AND Data[24]) AND (NOT Data[25])) AND (NOT Data[26]))) OR Data[30])) AND ((NOT ((((Data[21] AND Data[23]) AND Data[24]) AND (NOT Data[25])) AND (NOT Data[26]))) OR Data[31])) AND ((NOT (((((NOT Data[21]) AND (NOT Data[23])) AND (NOT Data[24])) AND Data[25]) AND (NOT Data[26]))) OR Data[22])) AND ((NOT ((((Data[21] AND (NOT Data[23])) AND (NOT Data[24])) AND Data[25]) AND (NOT Data[26]))) OR Data[33])) AND ((NOT (((((NOT Data[21]) AND Data[23]) AND (NOT Data[24])) AND Data[25]) AND (NOT Data[26]))) OR Data[9])) AND ((NOT ((((Data[21] AND Data[23]) AND (NOT Data[24])) AND Data[25]) AND (NOT Data[26]))) OR Data[32])) AND ((NOT (((((NOT Data[21]) AND (NOT Data[23])) AND Data[24]) AND Data[25]) AND (NOT Data[26]))) OR Data[28])) AND ((NOT ((((Data[21] AND (NOT Data[23])) AND Data[24]) AND Data[25]) AND (NOT Data[26]))) OR Data[34])) AND ((NOT (((((NOT Data[21]) AND Data[23]) AND Data[24]) AND Data[25]) AND (NOT Data[26]))) OR Data[37])) AND ((NOT ((((Data[21] AND Data[23]) AND Data[24]) AND Data[25]) AND (NOT Data[26]))) OR Data[2])) AND ((NOT (((((NOT Data[21]) AND (NOT Data[23])) AND (NOT Data[24])) AND (NOT Data[25])) AND Data[26])) OR Data[29])) AND ((NOT ((((Data[21] AND (NOT Data[23])) AND (NOT Data[24])) AND (NOT Data[25])) AND Data[26])) OR Data[36])) AND ((NOT (((((NOT Data[21]) AND Data[23]) AND (NOT Data[24])) AND (NOT Data[25])) AND Data[26])) OR Data[3])) AND ((NOT ((((Data[21] AND Data[23]) AND (NOT Data[24])) AND (NOT Data[25])) AND Data[26])) OR Data[7])) AND ((NOT (((((NOT Data[21]) AND (NOT Data[23])) AND Data[24]) AND (NOT Data[25])) AND Data[26])) OR Data[35])) AND ((NOT ((((Data[21] AND (NOT Data[23])) AND Data[24]) AND (NOT Data[25])) AND Data[26])) OR Data[8])) AND ((NOT (((((NOT Data[21]) AND Data[23]) AND Data[24]) AND (NOT Data[25])) AND Data[26])) OR Data[13])) AND ((NOT ((((Data[21] AND Data[23]) AND Data[24]) AND (NOT Data[25])) AND Data[26])) OR Data[12])) AND ((NOT (((((NOT Data[21]) AND (NOT Data[23])) AND (NOT Data[24])) AND Data[25]) AND Data[26])) OR Data[11])) AND ((NOT ((((Data[21] AND (NOT Data[23])) AND (NOT Data[24])) AND Data[25]) AND Data[26])) OR Data[19])) AND ((NOT (((((NOT Data[21]) AND Data[23]) AND (NOT Data[24])) AND Data[25]) AND Data[26])) OR Data[18])) AND ((NOT ((((Data[21] AND Data[23]) AND (NOT Data[24])) AND Data[25]) AND Data[26])) OR Data[15])) AND ((NOT (((((NOT Data[21]) AND (NOT Data[23])) AND Data[24]) AND Data[25]) AND Data[26])) OR Data[10])) AND ((NOT ((((Data[21] AND (NOT Data[23])) AND Data[24]) AND Data[25]) AND Data[26])) OR Data[14])) AND ((NOT (((((NOT Data[21]) AND Data[23]) AND Data[24]) AND Data[25]) AND Data[26])) OR Data[16])) AND ((NOT ((((Data[21] AND Data[23]) AND Data[24]) AND Data[25]) AND Data[26])) OR Data[17]));
    OutReady := 1;
    CollectInput(RESET:=TRUE);
  END_IF;
END_PROGRAM

CONFIGURATION Config0
  RESOURCE Res0 ON PLC
    TASK task0(INTERVAL := T#20ms,PRIORITY := 0);
    PROGRAM instance0 WITH task0 : Boiler;
  END_RESOURCE
END_CONFIGURATION

(* ---- 5-MUX_gloms-friar-gimme.st ---- *)
(*
This code implements a shuffled multiplexer with 5 control bits.
The control bits are: Data[N23], Data[N2], Data[N20], Data[N3], Data[N4]
The input bits are: Data[N21], Data[N26], Data[N1], Data[N22], Data[N25], Data[N24], Data[N5], Data[N6], Data[N31], Data[N33], Data[N8], Data[N27], Data[N30], Data[N29], Data[N9], Data[N32], Data[N12], Data[N10], Data[N28], Data[N7], Data[N13], Data[N14], Data[N11], Data[N34], Data[N35], Data[N37], Data[N15], Data[N16], Data[N36], Data[N17], Data[N18], Data[N19]

The symbolic expression is:
((((((((((((((((((((((((((((((((!(((((!(IN23)) & (!(IN2))) & (!(IN20))) & (!(IN3))) & (!(IN4)))) | IN21) & ((!((((IN23 & (!(IN2))) & (!(IN20))) & (!(IN3))) & (!(IN4)))) | IN26)) & ((!(((((!(IN23)) & IN2) & (!(IN20))) & (!(IN3))) & (!(IN4)))) | IN1)) & ((!((((IN23 & IN2) & (!(IN20))) & (!(IN3))) & (!(IN4)))) | IN22)) & ((!(((((!(IN23)) & (!(IN2))) & IN20) & (!(IN3))) & (!(IN4)))) | IN25)) & ((!((((IN23 & (!(IN2))) & IN20) & (!(IN3))) & (!(IN4)))) | IN24)) & ((!(((((!(IN23)) & IN2) & IN20) & (!(IN3))) & (!(IN4)))) | IN5)) & ((!((((IN23 & IN2) & IN20) & (!(IN3))) & (!(IN4)))) | IN6)) & ((!(((((!(IN23)) & (!(IN2))) & (!(IN20))) & IN3) & (!(IN4)))) | IN31)) & ((!((((IN23 & (!(IN2))) & (!(IN20))) & IN3) & (!(IN4)))) | IN33)) & ((!(((((!(IN23)) & IN2) & (!(IN20))) & IN3) & (!(IN4)))) | IN8)) & ((!((((IN23 & IN2) & (!(IN20))) & IN3) & (!(IN4)))) | IN27)) & ((!(((((!(IN23)) & (!(IN2))) & IN20) & IN3) & (!(IN4)))) | IN30)) & ((!((((IN23 & (!(IN2))) & IN20) & IN3) & (!(IN4)))) | IN29)) & ((!(((((!(IN23)) & IN2) & IN20) & IN3) & (!(IN4)))) | IN9)) & ((!((((IN23 & IN2) & IN20) & IN3) & (!(IN4)))) | IN32)) & ((!(((((!(IN23)) & (!(IN2))) & (!(IN20))) & (!(IN3))) & IN4)) | IN12)) & ((!((((IN23 & (!(IN2))) & (!(IN20))) & (!(IN3))) & IN4)) | IN10)) & ((!(((((!(IN23)) & IN2) & (!(IN20))) & (!(IN3))) & IN4)) | IN28)) & ((!((((IN23 & IN2) & (!(IN20))) & (!(IN3))) & IN4)) | IN7)) & ((!(((((!(IN23)) & (!(IN2))) & IN20) & (!(IN3))) & IN4)) | IN13)) & ((!((((IN23 & (!(IN2))) & IN20) & (!(IN3))) & IN4)) | IN14)) & ((!(((((!(IN23)) & IN2) & IN20) & (!(IN3))) & IN4)) | IN11)) & ((!((((IN23 & IN2) & IN20) & (!(IN3))) & IN4)) | IN34)) & ((!(((((!(IN23)) & (!(IN2))) & (!(IN20))) & IN3) & IN4)) | IN35)) & ((!((((IN23 & (!(IN2))) & (!(IN20))) & IN3) & IN4)) | IN37)) & ((!(((((!(IN23)) & IN2) & (!(IN20))) & IN3) & IN4)) | IN15)) & ((!((((IN23 & IN2) & (!(IN20))) & IN3) & IN4)) | IN16)) & ((!(((((!(IN23)) & (!(IN2))) & IN20) & IN3) & IN4)) | IN36)) & ((!((((IN23 & (!(IN2))) & IN20) & IN3) & IN4)) | IN17)) & ((!(((((!(IN23)) & IN2) & IN20) & IN3) & IN4)) | IN18)) & ((!((((IN23 & IN2) & IN20) & IN3) & IN4)) | IN19)

*)

FUNCTION_BLOCK F_CollectInput
  VAR_IN_OUT
      Data : ARRAY[1..40] OF BOOL;
  END_VAR
  VAR_INPUT
      TICK  : BOOL := 0;
      IN1   : BOOL := 0;
      IN2   : BOOL := 0;
      IN3   : BOOL := 0;
      IN4   : BOOL := 0;
      IN5   : BOOL := 0;
      RESET : BOOL := FALSE;
  END_VAR
  VAR_OUTPUT
      Finished : BOOL;
  END_VAR
  VAR
      j    : USINT := 1;
      tock : BOOL  := 0;
  END_VAR
  IF NOT RESET AND tock = NOT TICK THEN
      Data[j]   := IN1;
      Data[j+1] := IN2;
      Data[j+2] := IN3;
      Data[j+3] := IN4;
      Data[j+4] := IN5;
      j := j + 5;
      tock := TICK;
  ELSE
      j := 1;
      tock := 0;
  END_IF;
  Finished := (j > 40);
END_FUNCTION_BLOCK

PROGRAM Boiler
  VAR
    Data  : ARRAY[1..40] OF BOOL;
    Ready : BOOL;
    CollectInput : F_CollectInput;
  END_VAR
  VAR
    TICK     AT %IX1.0 : BOOL;
    IN1      AT %IX0.3 : BOOL;
    IN2      AT %IX0.4 : BOOL;
    IN3      AT %IX0.5 : BOOL;
    IN4      AT %IX0.6 : BOOL;
    IN5      AT %IX0.7 : BOOL;
    OutReady AT %QX0.0 : BOOL := FALSE;
    FeedNext AT %QX0.1 : BOOL := FALSE;
    Out      AT %QX0.2 : BOOL;
  END_VAR
  CollectInput(TICK:=TICK, IN1:=IN1, IN2:=IN2, IN3:=IN3, IN4:=IN4, IN5:=IN5);
  Ready := CollectInput.Finished;
  FeedNext := 1;
  IF Ready THEN
    Out := (((((((((((((((((((((((((((((((((NOT (((((NOT Data[23]) AND (NOT Data[2])) AND (NOT Data[20])) AND (NOT Data[3])) AND (NOT Data[4]))) OR Data[21]) AND ((NOT ((((Data[23] AND (NOT Data[2])) AND (NOT Data[20])) AND (NOT Data[3])) AND (NOT Data[4]))) OR Data[26])) AND ((NOT (((((NOT Data[23]) AND Data[2]) AND (NOT Data[20])) AND (NOT Data[3])) AND (NOT Data[4]))) OR Data[1])) AND ((NOT ((((Data[23] AND Data[2]) AND (NOT Data[20])) AND (NOT Data[3])) AND (NOT Data[4]))) OR Data[22])) AND ((NOT (((((NOT Data[23]) AND (NOT Data[2])) AND Data[20]) AND (NOT Data[3])) AND (NOT Data[4]))) OR Data[25])) AND ((NOT ((((Data[23] AND (NOT Data[2])) AND Data[20]) AND (NOT Data[3])) AND (NOT Data[4]))) OR Data[24])) AND ((NOT (((((NOT Data[23]) AND Data[2]) AND Data[20]) AND (NOT Data[3])) AND (NOT Data[4]))) OR Data[5])) AND ((NOT ((((Data[23] AND Data[2]) AND Data[20]) AND (NOT Data[3])) AND (NOT Data[4]))) OR Data[6])) AND ((NOT (((((NOT Data[23]) AND (NOT Data[2])) AND (NOT Data[20])) AND Data[3]) AND (NOT Data[4]))) OR Data[31])) AND ((NOT ((((Data[23] AND (NOT Data[2])) AND (NOT Data[20])) AND Data[3]) AND (NOT Data[4]))) OR Data[33])) AND ((NOT (((((NOT Data[23]) AND Data[2]) AND (NOT Data[20])) AND Data[3]) AND (NOT Data[4]))) OR Data[8])) AND ((NOT ((((Data[23] AND Data[2]) AND (NOT Data[20])) AND Data[3]) AND (NOT Data[4]))) OR Data[27])) AND ((NOT (((((NOT Data[23]) AND (NOT Data[2])) AND Data[20]) AND Data[3]) AND (NOT Data[4]))) OR Data[30])) AND ((NOT ((((Data[23] AND (NOT Data[2])) AND Data[20]) AND Data[3]) AND (NOT Data[4]))) OR Data[29])) AND ((NOT (((((NOT Data[23]) AND Data[2]) AND Data[20]) AND Data[3]) AND (NOT Data[4]))) OR Data[9])) AND ((NOT ((((Data[23] AND Data[2]) AND Data[20]) AND Data[3]) AND (NOT Data[4]))) OR Data[32])) AND ((NOT (((((NOT Data[23]) AND (NOT Data[2])) AND (NOT Data[20])) AND (NOT Data[3])) AND Data[4])) OR Data[12])) AND ((NOT ((((Data[23] AND (NOT Data[2])) AND (NOT Data[20])) AND (NOT Data[3])) AND Data[4])) OR Data[10])) AND ((NOT (((((NOT Data[23]) AND Data[2]) AND (NOT Data[20])) AND (NOT Data[3])) AND Data[4])) OR Data[28])) AND ((NOT ((((Data[23] AND Data[2]) AND (NOT Data[20])) AND (NOT Data[3])) AND Data[4])) OR Data[7])) AND ((NOT (((((NOT Data[23]) AND (NOT Data[2])) AND Data[20]) AND (NOT Data[3])) AND Data[4])) OR Data[13])) AND ((NOT ((((Data[23] AND (NOT Data[2])) AND Data[20]) AND (NOT Data[3])) AND Data[4])) OR Data[14])) AND ((NOT (((((NOT Data[23]) AND Data[2]) AND Data[20]) AND (NOT Data[3])) AND Data[4])) OR Data[11])) AND ((NOT ((((Data[23] AND Data[2]) AND Data[20]) AND (NOT Data[3])) AND Data[4])) OR Data[34])) AND ((NOT (((((NOT Data[23]) AND (NOT Data[2])) AND (NOT Data[20])) AND Data[3]) AND Data[4])) OR Data[35])) AND ((NOT ((((Data[23] AND (NOT Data[2])) AND (NOT Data[20])) AND Data[3]) AND Data[4])) OR Data[37])) AND ((NOT (((((NOT Data[23]) AND Data[2]) AND (NOT Data[20])) AND Data[3]) AND Data[4])) OR Data[15])) AND ((NOT ((((Data[23] AND Data[2]) AND (NOT Data[20])) AND Data[3]) AND Data[4])) OR Data[16])) AND ((NOT (((((NOT Data[23]) AND (NOT Data[2])) AND Data[20]) AND Data[3]) AND Data[4])) OR Data[36])) AND ((NOT ((((Data[23] AND (NOT Data[2])) AND Data[20]) AND Data[3]) AND Data[4])) OR Data[17])) AND ((NOT (((((NOT Data[23]) AND Data[2]) AND Data[20]) AND Data[3]) AND Data[4])) OR Data[18])) AND ((NOT ((((Data[23] AND Data[2]) AND Data[20]) AND Data[3]) AND Data[4])) OR Data[19]));
    OutReady := 1;
    CollectInput(RESET:=TRUE);
  END_IF;
END_PROGRAM

CONFIGURATION Config0
  RESOURCE Res0 ON PLC
    TASK task0(INTERVAL := T#20ms,PRIORITY := 0);
    PROGRAM instance0 WITH task0 : Boiler;
  END_RESOURCE
END_CONFIGURATION

(* ---- 5-MUX_gluts-trial-bevel.st ---- *)
(*
This code implements a shuffled multiplexer with 5 control bits.
The control bits are: Data[N23], Data[N3], Data[N2], Data[N1], Data[N21]
The input bits are: Data[N20], Data[N24], Data[N22], Data[N4], Data[N25], Data[N26], Data[N27], Data[N6], Data[N31], Data[N5], Data[N7], Data[N28], Data[N30], Data[N29], Data[N35], Data[N32], Data[N33], Data[N34], Data[N9], Data[N36], Data[N37], Data[N8], Data[N10], Data[N13], Data[N11], Data[N12], Data[N15], Data[N14], Data[N17], Data[N16], Data[N18], Data[N19]

The symbolic expression is:
((((((((((((((((((((((((((((((((!(((((!(IN23)) & (!(IN3))) & (!(IN2))) & (!(IN1))) & (!(IN21)))) | IN20) & ((!((((IN23 & (!(IN3))) & (!(IN2))) & (!(IN1))) & (!(IN21)))) | IN24)) & ((!(((((!(IN23)) & IN3) & (!(IN2))) & (!(IN1))) & (!(IN21)))) | IN22)) & ((!((((IN23 & IN3) & (!(IN2))) & (!(IN1))) & (!(IN21)))) | IN4)) & ((!(((((!(IN23)) & (!(IN3))) & IN2) & (!(IN1))) & (!(IN21)))) | IN25)) & ((!((((IN23 & (!(IN3))) & IN2) & (!(IN1))) & (!(IN21)))) | IN26)) & ((!(((((!(IN23)) & IN3) & IN2) & (!(IN1))) & (!(IN21)))) | IN27)) & ((!((((IN23 & IN3) & IN2) & (!(IN1))) & (!(IN21)))) | IN6)) & ((!(((((!(IN23)) & (!(IN3))) & (!(IN2))) & IN1) & (!(IN21)))) | IN31)) & ((!((((IN23 & (!(IN3))) & (!(IN2))) & IN1) & (!(IN21)))) | IN5)) & ((!(((((!(IN23)) & IN3) & (!(IN2))) & IN1) & (!(IN21)))) | IN7)) & ((!((((IN23 & IN3) & (!(IN2))) & IN1) & (!(IN21)))) | IN28)) & ((!(((((!(IN23)) & (!(IN3))) & IN2) & IN1) & (!(IN21)))) | IN30)) & ((!((((IN23 & (!(IN3))) & IN2) & IN1) & (!(IN21)))) | IN29)) & ((!(((((!(IN23)) & IN3) & IN2) & IN1) & (!(IN21)))) | IN35)) & ((!((((IN23 & IN3) & IN2) & IN1) & (!(IN21)))) | IN32)) & ((!(((((!(IN23)) & (!(IN3))) & (!(IN2))) & (!(IN1))) & IN21)) | IN33)) & ((!((((IN23 & (!(IN3))) & (!(IN2))) & (!(IN1))) & IN21)) | IN34)) & ((!(((((!(IN23)) & IN3) & (!(IN2))) & (!(IN1))) & IN21)) | IN9)) & ((!((((IN23 & IN3) & (!(IN2))) & (!(IN1))) & IN21)) | IN36)) & ((!(((((!(IN23)) & (!(IN3))) & IN2) & (!(IN1))) & IN21)) | IN37)) & ((!((((IN23 & (!(IN3))) & IN2) & (!(IN1))) & IN21)) | IN8)) & ((!(((((!(IN23)) & IN3) & IN2) & (!(IN1))) & IN21)) | IN10)) & ((!((((IN23 & IN3) & IN2) & (!(IN1))) & IN21)) | IN13)) & ((!(((((!(IN23)) & (!(IN3))) & (!(IN2))) & IN1) & IN21)) | IN11)) & ((!((((IN23 & (!(IN3))) & (!(IN2))) & IN1) & IN21)) | IN12)) & ((!(((((!(IN23)) & IN3) & (!(IN2))) & IN1) & IN21)) | IN15)) & ((!((((IN23 & IN3) & (!(IN2))) & IN1) & IN21)) | IN14)) & ((!(((((!(IN23)) & (!(IN3))) & IN2) & IN1) & IN21)) | IN17)) & ((!((((IN23 & (!(IN3))) & IN2) & IN1) & IN21)) | IN16)) & ((!(((((!(IN23)) & IN3) & IN2) & IN1) & IN21)) | IN18)) & ((!((((IN23 & IN3) & IN2) & IN1) & IN21)) | IN19)

*)

FUNCTION_BLOCK F_CollectInput
  VAR_IN_OUT
      Data : ARRAY[1..40] OF BOOL;
  END_VAR
  VAR_INPUT
      TICK  : BOOL := 0;
      IN1   : BOOL := 0;
      IN2   : BOOL := 0;
      IN3   : BOOL := 0;
      IN4   : BOOL := 0;
      IN5   : BOOL := 0;
      RESET : BOOL := FALSE;
  END_VAR
  VAR_OUTPUT
      Finished : BOOL;
  END_VAR
  VAR
      j    : USINT := 1;
      tock : BOOL  := 0;
  END_VAR
  IF NOT RESET AND tock = NOT TICK THEN
      Data[j]   := IN1;
      Data[j+1] := IN2;
      Data[j+2] := IN3;
      Data[j+3] := IN4;
      Data[j+4] := IN5;
      j := j + 5;
      tock := TICK;
  ELSE
      j := 1;
      tock := 0;
  END_IF;
  Finished := (j > 40);
END_FUNCTION_BLOCK

PROGRAM Boiler
  VAR
    Data  : ARRAY[1..40] OF BOOL;
    Ready : BOOL;
    CollectInput : F_CollectInput;
  END_VAR
  VAR
    TICK     AT %IX1.0 : BOOL;
    IN1      AT %IX0.3 : BOOL;
    IN2      AT %IX0.4 : BOOL;
    IN3      AT %IX0.5 : BOOL;
    IN4      AT %IX0.6 : BOOL;
    IN5      AT %IX0.7 : BOOL;
    OutReady AT %QX0.0 : BOOL := FALSE;
    FeedNext AT %QX0.1 : BOOL := FALSE;
    Out      AT %QX0.2 : BOOL;
  END_VAR
  CollectInput(TICK:=TICK, IN1:=IN1, IN2:=IN2, IN3:=IN3, IN4:=IN4, IN5:=IN5);
  Ready := CollectInput.Finished;
  FeedNext := 1;
  IF Ready THEN
    Out := (((((((((((((((((((((((((((((((((NOT (((((NOT Data[23]) AND (NOT Data[3])) AND (NOT Data[2])) AND (NOT Data[1])) AND (NOT Data[21]))) OR Data[20]) AND ((NOT ((((Data[23] AND (NOT Data[3])) AND (NOT Data[2])) AND (NOT Data[1])) AND (NOT Data[21]))) OR Data[24])) AND ((NOT (((((NOT Data[23]) AND Data[3]) AND (NOT Data[2])) AND (NOT Data[1])) AND (NOT Data[21]))) OR Data[22])) AND ((NOT ((((Data[23] AND Data[3]) AND (NOT Data[2])) AND (NOT Data[1])) AND (NOT Data[21]))) OR Data[4])) AND ((NOT (((((NOT Data[23]) AND (NOT Data[3])) AND Data[2]) AND (NOT Data[1])) AND (NOT Data[21]))) OR Data[25])) AND ((NOT ((((Data[23] AND (NOT Data[3])) AND Data[2]) AND (NOT Data[1])) AND (NOT Data[21]))) OR Data[26])) AND ((NOT (((((NOT Data[23]) AND Data[3]) AND Data[2]) AND (NOT Data[1])) AND (NOT Data[21]))) OR Data[27])) AND ((NOT ((((Data[23] AND Data[3]) AND Data[2]) AND (NOT Data[1])) AND (NOT Data[21]))) OR Data[6])) AND ((NOT (((((NOT Data[23]) AND (NOT Data[3])) AND (NOT Data[2])) AND Data[1]) AND (NOT Data[21]))) OR Data[31])) AND ((NOT ((((Data[23] AND (NOT Data[3])) AND (NOT Data[2])) AND Data[1]) AND (NOT Data[21]))) OR Data[5])) AND ((NOT (((((NOT Data[23]) AND Data[3]) AND (NOT Data[2])) AND Data[1]) AND (NOT Data[21]))) OR Data[7])) AND ((NOT ((((Data[23] AND Data[3]) AND (NOT Data[2])) AND Data[1]) AND (NOT Data[21]))) OR Data[28])) AND ((NOT (((((NOT Data[23]) AND (NOT Data[3])) AND Data[2]) AND Data[1]) AND (NOT Data[21]))) OR Data[30])) AND ((NOT ((((Data[23] AND (NOT Data[3])) AND Data[2]) AND Data[1]) AND (NOT Data[21]))) OR Data[29])) AND ((NOT (((((NOT Data[23]) AND Data[3]) AND Data[2]) AND Data[1]) AND (NOT Data[21]))) OR Data[35])) AND ((NOT ((((Data[23] AND Data[3]) AND Data[2]) AND Data[1]) AND (NOT Data[21]))) OR Data[32])) AND ((NOT (((((NOT Data[23]) AND (NOT Data[3])) AND (NOT Data[2])) AND (NOT Data[1])) AND Data[21])) OR Data[33])) AND ((NOT ((((Data[23] AND (NOT Data[3])) AND (NOT Data[2])) AND (NOT Data[1])) AND Data[21])) OR Data[34])) AND ((NOT (((((NOT Data[23]) AND Data[3]) AND (NOT Data[2])) AND (NOT Data[1])) AND Data[21])) OR Data[9])) AND ((NOT ((((Data[23] AND Data[3]) AND (NOT Data[2])) AND (NOT Data[1])) AND Data[21])) OR Data[36])) AND ((NOT (((((NOT Data[23]) AND (NOT Data[3])) AND Data[2]) AND (NOT Data[1])) AND Data[21])) OR Data[37])) AND ((NOT ((((Data[23] AND (NOT Data[3])) AND Data[2]) AND (NOT Data[1])) AND Data[21])) OR Data[8])) AND ((NOT (((((NOT Data[23]) AND Data[3]) AND Data[2]) AND (NOT Data[1])) AND Data[21])) OR Data[10])) AND ((NOT ((((Data[23] AND Data[3]) AND Data[2]) AND (NOT Data[1])) AND Data[21])) OR Data[13])) AND ((NOT (((((NOT Data[23]) AND (NOT Data[3])) AND (NOT Data[2])) AND Data[1]) AND Data[21])) OR Data[11])) AND ((NOT ((((Data[23] AND (NOT Data[3])) AND (NOT Data[2])) AND Data[1]) AND Data[21])) OR Data[12])) AND ((NOT (((((NOT Data[23]) AND Data[3]) AND (NOT Data[2])) AND Data[1]) AND Data[21])) OR Data[15])) AND ((NOT ((((Data[23] AND Data[3]) AND (NOT Data[2])) AND Data[1]) AND Data[21])) OR Data[14])) AND ((NOT (((((NOT Data[23]) AND (NOT Data[3])) AND Data[2]) AND Data[1]) AND Data[21])) OR Data[17])) AND ((NOT ((((Data[23] AND (NOT Data[3])) AND Data[2]) AND Data[1]) AND Data[21])) OR Data[16])) AND ((NOT (((((NOT Data[23]) AND Data[3]) AND Data[2]) AND Data[1]) AND Data[21])) OR Data[18])) AND ((NOT ((((Data[23] AND Data[3]) AND Data[2]) AND Data[1]) AND Data[21])) OR Data[19]));
    OutReady := 1;
    CollectInput(RESET:=TRUE);
  END_IF;
END_PROGRAM

CONFIGURATION Config0
  RESOURCE Res0 ON PLC
    TASK task0(INTERVAL := T#20ms,PRIORITY := 0);
    PROGRAM instance0 WITH task0 : Boiler;
  END_RESOURCE
END_CONFIGURATION

(* ---- 5-MUX_gwine-knobs-await.st ---- *)
(*
This code implements a shuffled multiplexer with 5 control bits.
The control bits are: Data[N22], Data[N3], Data[N2], Data[N20], Data[N4]
The input bits are: Data[N21], Data[N1], Data[N6], Data[N5], Data[N26], Data[N9], Data[N23], Data[N24], Data[N8], Data[N25], Data[N7], Data[N27], Data[N11], Data[N12], Data[N28], Data[N31], Data[N10], Data[N13], Data[N29], Data[N30], Data[N15], Data[N33], Data[N14], Data[N32], Data[N35], Data[N18], Data[N17], Data[N37], Data[N16], Data[N34], Data[N36], Data[N19]

The symbolic expression is:
((((((((((((((((((((((((((((((((!(((((!(IN22)) & (!(IN3))) & (!(IN2))) & (!(IN20))) & (!(IN4)))) | IN21) & ((!((((IN22 & (!(IN3))) & (!(IN2))) & (!(IN20))) & (!(IN4)))) | IN1)) & ((!(((((!(IN22)) & IN3) & (!(IN2))) & (!(IN20))) & (!(IN4)))) | IN6)) & ((!((((IN22 & IN3) & (!(IN2))) & (!(IN20))) & (!(IN4)))) | IN5)) & ((!(((((!(IN22)) & (!(IN3))) & IN2) & (!(IN20))) & (!(IN4)))) | IN26)) & ((!((((IN22 & (!(IN3))) & IN2) & (!(IN20))) & (!(IN4)))) | IN9)) & ((!(((((!(IN22)) & IN3) & IN2) & (!(IN20))) & (!(IN4)))) | IN23)) & ((!((((IN22 & IN3) & IN2) & (!(IN20))) & (!(IN4)))) | IN24)) & ((!(((((!(IN22)) & (!(IN3))) & (!(IN2))) & IN20) & (!(IN4)))) | IN8)) & ((!((((IN22 & (!(IN3))) & (!(IN2))) & IN20) & (!(IN4)))) | IN25)) & ((!(((((!(IN22)) & IN3) & (!(IN2))) & IN20) & (!(IN4)))) | IN7)) & ((!((((IN22 & IN3) & (!(IN2))) & IN20) & (!(IN4)))) | IN27)) & ((!(((((!(IN22)) & (!(IN3))) & IN2) & IN20) & (!(IN4)))) | IN11)) & ((!((((IN22 & (!(IN3))) & IN2) & IN20) & (!(IN4)))) | IN12)) & ((!(((((!(IN22)) & IN3) & IN2) & IN20) & (!(IN4)))) | IN28)) & ((!((((IN22 & IN3) & IN2) & IN20) & (!(IN4)))) | IN31)) & ((!(((((!(IN22)) & (!(IN3))) & (!(IN2))) & (!(IN20))) & IN4)) | IN10)) & ((!((((IN22 & (!(IN3))) & (!(IN2))) & (!(IN20))) & IN4)) | IN13)) & ((!(((((!(IN22)) & IN3) & (!(IN2))) & (!(IN20))) & IN4)) | IN29)) & ((!((((IN22 & IN3) & (!(IN2))) & (!(IN20))) & IN4)) | IN30)) & ((!(((((!(IN22)) & (!(IN3))) & IN2) & (!(IN20))) & IN4)) | IN15)) & ((!((((IN22 & (!(IN3))) & IN2) & (!(IN20))) & IN4)) | IN33)) & ((!(((((!(IN22)) & IN3) & IN2) & (!(IN20))) & IN4)) | IN14)) & ((!((((IN22 & IN3) & IN2) & (!(IN20))) & IN4)) | IN32)) & ((!(((((!(IN22)) & (!(IN3))) & (!(IN2))) & IN20) & IN4)) | IN35)) & ((!((((IN22 & (!(IN3))) & (!(IN2))) & IN20) & IN4)) | IN18)) & ((!(((((!(IN22)) & IN3) & (!(IN2))) & IN20) & IN4)) | IN17)) & ((!((((IN22 & IN3) & (!(IN2))) & IN20) & IN4)) | IN37)) & ((!(((((!(IN22)) & (!(IN3))) & IN2) & IN20) & IN4)) | IN16)) & ((!((((IN22 & (!(IN3))) & IN2) & IN20) & IN4)) | IN34)) & ((!(((((!(IN22)) & IN3) & IN2) & IN20) & IN4)) | IN36)) & ((!((((IN22 & IN3) & IN2) & IN20) & IN4)) | IN19)

*)

FUNCTION_BLOCK F_CollectInput
  VAR_IN_OUT
      Data : ARRAY[1..40] OF BOOL;
  END_VAR
  VAR_INPUT
      TICK  : BOOL := 0;
      IN1   : BOOL := 0;
      IN2   : BOOL := 0;
      IN3   : BOOL := 0;
      IN4   : BOOL := 0;
      IN5   : BOOL := 0;
      RESET : BOOL := FALSE;
  END_VAR
  VAR_OUTPUT
      Finished : BOOL;
  END_VAR
  VAR
      j    : USINT := 1;
      tock : BOOL  := 0;
  END_VAR
  IF NOT RESET AND tock = NOT TICK THEN
      Data[j]   := IN1;
      Data[j+1] := IN2;
      Data[j+2] := IN3;
      Data[j+3] := IN4;
      Data[j+4] := IN5;
      j := j + 5;
      tock := TICK;
  ELSE
      j := 1;
      tock := 0;
  END_IF;
  Finished := (j > 40);
END_FUNCTION_BLOCK

PROGRAM Boiler
  VAR
    Data  : ARRAY[1..40] OF BOOL;
    Ready : BOOL;
    CollectInput : F_CollectInput;
  END_VAR
  VAR
    TICK     AT %IX1.0 : BOOL;
    IN1      AT %IX0.3 : BOOL;
    IN2      AT %IX0.4 : BOOL;
    IN3      AT %IX0.5 : BOOL;
    IN4      AT %IX0.6 : BOOL;
    IN5      AT %IX0.7 : BOOL;
    OutReady AT %QX0.0 : BOOL := FALSE;
    FeedNext AT %QX0.1 : BOOL := FALSE;
    Out      AT %QX0.2 : BOOL;
  END_VAR
  CollectInput(TICK:=TICK, IN1:=IN1, IN2:=IN2, IN3:=IN3, IN4:=IN4, IN5:=IN5);
  Ready := CollectInput.Finished;
  FeedNext := 1;
  IF Ready THEN
    Out := (((((((((((((((((((((((((((((((((NOT (((((NOT Data[22]) AND (NOT Data[3])) AND (NOT Data[2])) AND (NOT Data[20])) AND (NOT Data[4]))) OR Data[21]) AND ((NOT ((((Data[22] AND (NOT Data[3])) AND (NOT Data[2])) AND (NOT Data[20])) AND (NOT Data[4]))) OR Data[1])) AND ((NOT (((((NOT Data[22]) AND Data[3]) AND (NOT Data[2])) AND (NOT Data[20])) AND (NOT Data[4]))) OR Data[6])) AND ((NOT ((((Data[22] AND Data[3]) AND (NOT Data[2])) AND (NOT Data[20])) AND (NOT Data[4]))) OR Data[5])) AND ((NOT (((((NOT Data[22]) AND (NOT Data[3])) AND Data[2]) AND (NOT Data[20])) AND (NOT Data[4]))) OR Data[26])) AND ((NOT ((((Data[22] AND (NOT Data[3])) AND Data[2]) AND (NOT Data[20])) AND (NOT Data[4]))) OR Data[9])) AND ((NOT (((((NOT Data[22]) AND Data[3]) AND Data[2]) AND (NOT Data[20])) AND (NOT Data[4]))) OR Data[23])) AND ((NOT ((((Data[22] AND Data[3]) AND Data[2]) AND (NOT Data[20])) AND (NOT Data[4]))) OR Data[24])) AND ((NOT (((((NOT Data[22]) AND (NOT Data[3])) AND (NOT Data[2])) AND Data[20]) AND (NOT Data[4]))) OR Data[8])) AND ((NOT ((((Data[22] AND (NOT Data[3])) AND (NOT Data[2])) AND Data[20]) AND (NOT Data[4]))) OR Data[25])) AND ((NOT (((((NOT Data[22]) AND Data[3]) AND (NOT Data[2])) AND Data[20]) AND (NOT Data[4]))) OR Data[7])) AND ((NOT ((((Data[22] AND Data[3]) AND (NOT Data[2])) AND Data[20]) AND (NOT Data[4]))) OR Data[27])) AND ((NOT (((((NOT Data[22]) AND (NOT Data[3])) AND Data[2]) AND Data[20]) AND (NOT Data[4]))) OR Data[11])) AND ((NOT ((((Data[22] AND (NOT Data[3])) AND Data[2]) AND Data[20]) AND (NOT Data[4]))) OR Data[12])) AND ((NOT (((((NOT Data[22]) AND Data[3]) AND Data[2]) AND Data[20]) AND (NOT Data[4]))) OR Data[28])) AND ((NOT ((((Data[22] AND Data[3]) AND Data[2]) AND Data[20]) AND (NOT Data[4]))) OR Data[31])) AND ((NOT (((((NOT Data[22]) AND (NOT Data[3])) AND (NOT Data[2])) AND (NOT Data[20])) AND Data[4])) OR Data[10])) AND ((NOT ((((Data[22] AND (NOT Data[3])) AND (NOT Data[2])) AND (NOT Data[20])) AND Data[4])) OR Data[13])) AND ((NOT (((((NOT Data[22]) AND Data[3]) AND (NOT Data[2])) AND (NOT Data[20])) AND Data[4])) OR Data[29])) AND ((NOT ((((Data[22] AND Data[3]) AND (NOT Data[2])) AND (NOT Data[20])) AND Data[4])) OR Data[30])) AND ((NOT (((((NOT Data[22]) AND (NOT Data[3])) AND Data[2]) AND (NOT Data[20])) AND Data[4])) OR Data[15])) AND ((NOT ((((Data[22] AND (NOT Data[3])) AND Data[2]) AND (NOT Data[20])) AND Data[4])) OR Data[33])) AND ((NOT (((((NOT Data[22]) AND Data[3]) AND Data[2]) AND (NOT Data[20])) AND Data[4])) OR Data[14])) AND ((NOT ((((Data[22] AND Data[3]) AND Data[2]) AND (NOT Data[20])) AND Data[4])) OR Data[32])) AND ((NOT (((((NOT Data[22]) AND (NOT Data[3])) AND (NOT Data[2])) AND Data[20]) AND Data[4])) OR Data[35])) AND ((NOT ((((Data[22] AND (NOT Data[3])) AND (NOT Data[2])) AND Data[20]) AND Data[4])) OR Data[18])) AND ((NOT (((((NOT Data[22]) AND Data[3]) AND (NOT Data[2])) AND Data[20]) AND Data[4])) OR Data[17])) AND ((NOT ((((Data[22] AND Data[3]) AND (NOT Data[2])) AND Data[20]) AND Data[4])) OR Data[37])) AND ((NOT (((((NOT Data[22]) AND (NOT Data[3])) AND Data[2]) AND Data[20]) AND Data[4])) OR Data[16])) AND ((NOT ((((Data[22] AND (NOT Data[3])) AND Data[2]) AND Data[20]) AND Data[4])) OR Data[34])) AND ((NOT (((((NOT Data[22]) AND Data[3]) AND Data[2]) AND Data[20]) AND Data[4])) OR Data[36])) AND ((NOT ((((Data[22] AND Data[3]) AND Data[2]) AND Data[20]) AND Data[4])) OR Data[19]));
    OutReady := 1;
    CollectInput(RESET:=TRUE);
  END_IF;
END_PROGRAM

CONFIGURATION Config0
  RESOURCE Res0 ON PLC
    TASK task0(INTERVAL := T#20ms,PRIORITY := 0);
    PROGRAM instance0 WITH task0 : Boiler;
  END_RESOURCE
END_CONFIGURATION

(* ---- 5-MUX_habit-loved-parry.st ---- *)
(*
This code implements a shuffled multiplexer with 5 control bits.
The control bits are: Data[N21], Data[N20], Data[N1], Data[N3], Data[N2]
The input bits are: Data[N26], Data[N4], Data[N24], Data[N25], Data[N6], Data[N22], Data[N23], Data[N27], Data[N28], Data[N31], Data[N29], Data[N30], Data[N5], Data[N8], Data[N37], Data[N9], Data[N32], Data[N35], Data[N33], Data[N7], Data[N10], Data[N11], Data[N36], Data[N12], Data[N13], Data[N15], Data[N16], Data[N34], Data[N14], Data[N17], Data[N18], Data[N19]

The symbolic expression is:
((((((((((((((((((((((((((((((((!(((((!(IN21)) & (!(IN20))) & (!(IN1))) & (!(IN3))) & (!(IN2)))) | IN26) & ((!((((IN21 & (!(IN20))) & (!(IN1))) & (!(IN3))) & (!(IN2)))) | IN4)) & ((!(((((!(IN21)) & IN20) & (!(IN1))) & (!(IN3))) & (!(IN2)))) | IN24)) & ((!((((IN21 & IN20) & (!(IN1))) & (!(IN3))) & (!(IN2)))) | IN25)) & ((!(((((!(IN21)) & (!(IN20))) & IN1) & (!(IN3))) & (!(IN2)))) | IN6)) & ((!((((IN21 & (!(IN20))) & IN1) & (!(IN3))) & (!(IN2)))) | IN22)) & ((!(((((!(IN21)) & IN20) & IN1) & (!(IN3))) & (!(IN2)))) | IN23)) & ((!((((IN21 & IN20) & IN1) & (!(IN3))) & (!(IN2)))) | IN27)) & ((!(((((!(IN21)) & (!(IN20))) & (!(IN1))) & IN3) & (!(IN2)))) | IN28)) & ((!((((IN21 & (!(IN20))) & (!(IN1))) & IN3) & (!(IN2)))) | IN31)) & ((!(((((!(IN21)) & IN20) & (!(IN1))) & IN3) & (!(IN2)))) | IN29)) & ((!((((IN21 & IN20) & (!(IN1))) & IN3) & (!(IN2)))) | IN30)) & ((!(((((!(IN21)) & (!(IN20))) & IN1) & IN3) & (!(IN2)))) | IN5)) & ((!((((IN21 & (!(IN20))) & IN1) & IN3) & (!(IN2)))) | IN8)) & ((!(((((!(IN21)) & IN20) & IN1) & IN3) & (!(IN2)))) | IN37)) & ((!((((IN21 & IN20) & IN1) & IN3) & (!(IN2)))) | IN9)) & ((!(((((!(IN21)) & (!(IN20))) & (!(IN1))) & (!(IN3))) & IN2)) | IN32)) & ((!((((IN21 & (!(IN20))) & (!(IN1))) & (!(IN3))) & IN2)) | IN35)) & ((!(((((!(IN21)) & IN20) & (!(IN1))) & (!(IN3))) & IN2)) | IN33)) & ((!((((IN21 & IN20) & (!(IN1))) & (!(IN3))) & IN2)) | IN7)) & ((!(((((!(IN21)) & (!(IN20))) & IN1) & (!(IN3))) & IN2)) | IN10)) & ((!((((IN21 & (!(IN20))) & IN1) & (!(IN3))) & IN2)) | IN11)) & ((!(((((!(IN21)) & IN20) & IN1) & (!(IN3))) & IN2)) | IN36)) & ((!((((IN21 & IN20) & IN1) & (!(IN3))) & IN2)) | IN12)) & ((!(((((!(IN21)) & (!(IN20))) & (!(IN1))) & IN3) & IN2)) | IN13)) & ((!((((IN21 & (!(IN20))) & (!(IN1))) & IN3) & IN2)) | IN15)) & ((!(((((!(IN21)) & IN20) & (!(IN1))) & IN3) & IN2)) | IN16)) & ((!((((IN21 & IN20) & (!(IN1))) & IN3) & IN2)) | IN34)) & ((!(((((!(IN21)) & (!(IN20))) & IN1) & IN3) & IN2)) | IN14)) & ((!((((IN21 & (!(IN20))) & IN1) & IN3) & IN2)) | IN17)) & ((!(((((!(IN21)) & IN20) & IN1) & IN3) & IN2)) | IN18)) & ((!((((IN21 & IN20) & IN1) & IN3) & IN2)) | IN19)

*)

FUNCTION_BLOCK F_CollectInput
  VAR_IN_OUT
      Data : ARRAY[1..40] OF BOOL;
  END_VAR
  VAR_INPUT
      TICK  : BOOL := 0;
      IN1   : BOOL := 0;
      IN2   : BOOL := 0;
      IN3   : BOOL := 0;
      IN4   : BOOL := 0;
      IN5   : BOOL := 0;
      RESET : BOOL := FALSE;
  END_VAR
  VAR_OUTPUT
      Finished : BOOL;
  END_VAR
  VAR
      j    : USINT := 1;
      tock : BOOL  := 0;
  END_VAR
  IF NOT RESET AND tock = NOT TICK THEN
      Data[j]   := IN1;
      Data[j+1] := IN2;
      Data[j+2] := IN3;
      Data[j+3] := IN4;
      Data[j+4] := IN5;
      j := j + 5;
      tock := TICK;
  ELSE
      j := 1;
      tock := 0;
  END_IF;
  Finished := (j > 40);
END_FUNCTION_BLOCK

PROGRAM Boiler
  VAR
    Data  : ARRAY[1..40] OF BOOL;
    Ready : BOOL;
    CollectInput : F_CollectInput;
  END_VAR
  VAR
    TICK     AT %IX1.0 : BOOL;
    IN1      AT %IX0.3 : BOOL;
    IN2      AT %IX0.4 : BOOL;
    IN3      AT %IX0.5 : BOOL;
    IN4      AT %IX0.6 : BOOL;
    IN5      AT %IX0.7 : BOOL;
    OutReady AT %QX0.0 : BOOL := FALSE;
    FeedNext AT %QX0.1 : BOOL := FALSE;
    Out      AT %QX0.2 : BOOL;
  END_VAR
  CollectInput(TICK:=TICK, IN1:=IN1, IN2:=IN2, IN3:=IN3, IN4:=IN4, IN5:=IN5);
  Ready := CollectInput.Finished;
  FeedNext := 1;
  IF Ready THEN
    Out := (((((((((((((((((((((((((((((((((NOT (((((NOT Data[21]) AND (NOT Data[20])) AND (NOT Data[1])) AND (NOT Data[3])) AND (NOT Data[2]))) OR Data[26]) AND ((NOT ((((Data[21] AND (NOT Data[20])) AND (NOT Data[1])) AND (NOT Data[3])) AND (NOT Data[2]))) OR Data[4])) AND ((NOT (((((NOT Data[21]) AND Data[20]) AND (NOT Data[1])) AND (NOT Data[3])) AND (NOT Data[2]))) OR Data[24])) AND ((NOT ((((Data[21] AND Data[20]) AND (NOT Data[1])) AND (NOT Data[3])) AND (NOT Data[2]))) OR Data[25])) AND ((NOT (((((NOT Data[21]) AND (NOT Data[20])) AND Data[1]) AND (NOT Data[3])) AND (NOT Data[2]))) OR Data[6])) AND ((NOT ((((Data[21] AND (NOT Data[20])) AND Data[1]) AND (NOT Data[3])) AND (NOT Data[2]))) OR Data[22])) AND ((NOT (((((NOT Data[21]) AND Data[20]) AND Data[1]) AND (NOT Data[3])) AND (NOT Data[2]))) OR Data[23])) AND ((NOT ((((Data[21] AND Data[20]) AND Data[1]) AND (NOT Data[3])) AND (NOT Data[2]))) OR Data[27])) AND ((NOT (((((NOT Data[21]) AND (NOT Data[20])) AND (NOT Data[1])) AND Data[3]) AND (NOT Data[2]))) OR Data[28])) AND ((NOT ((((Data[21] AND (NOT Data[20])) AND (NOT Data[1])) AND Data[3]) AND (NOT Data[2]))) OR Data[31])) AND ((NOT (((((NOT Data[21]) AND Data[20]) AND (NOT Data[1])) AND Data[3]) AND (NOT Data[2]))) OR Data[29])) AND ((NOT ((((Data[21] AND Data[20]) AND (NOT Data[1])) AND Data[3]) AND (NOT Data[2]))) OR Data[30])) AND ((NOT (((((NOT Data[21]) AND (NOT Data[20])) AND Data[1]) AND Data[3]) AND (NOT Data[2]))) OR Data[5])) AND ((NOT ((((Data[21] AND (NOT Data[20])) AND Data[1]) AND Data[3]) AND (NOT Data[2]))) OR Data[8])) AND ((NOT (((((NOT Data[21]) AND Data[20]) AND Data[1]) AND Data[3]) AND (NOT Data[2]))) OR Data[37])) AND ((NOT ((((Data[21] AND Data[20]) AND Data[1]) AND Data[3]) AND (NOT Data[2]))) OR Data[9])) AND ((NOT (((((NOT Data[21]) AND (NOT Data[20])) AND (NOT Data[1])) AND (NOT Data[3])) AND Data[2])) OR Data[32])) AND ((NOT ((((Data[21] AND (NOT Data[20])) AND (NOT Data[1])) AND (NOT Data[3])) AND Data[2])) OR Data[35])) AND ((NOT (((((NOT Data[21]) AND Data[20]) AND (NOT Data[1])) AND (NOT Data[3])) AND Data[2])) OR Data[33])) AND ((NOT ((((Data[21] AND Data[20]) AND (NOT Data[1])) AND (NOT Data[3])) AND Data[2])) OR Data[7])) AND ((NOT (((((NOT Data[21]) AND (NOT Data[20])) AND Data[1]) AND (NOT Data[3])) AND Data[2])) OR Data[10])) AND ((NOT ((((Data[21] AND (NOT Data[20])) AND Data[1]) AND (NOT Data[3])) AND Data[2])) OR Data[11])) AND ((NOT (((((NOT Data[21]) AND Data[20]) AND Data[1]) AND (NOT Data[3])) AND Data[2])) OR Data[36])) AND ((NOT ((((Data[21] AND Data[20]) AND Data[1]) AND (NOT Data[3])) AND Data[2])) OR Data[12])) AND ((NOT (((((NOT Data[21]) AND (NOT Data[20])) AND (NOT Data[1])) AND Data[3]) AND Data[2])) OR Data[13])) AND ((NOT ((((Data[21] AND (NOT Data[20])) AND (NOT Data[1])) AND Data[3]) AND Data[2])) OR Data[15])) AND ((NOT (((((NOT Data[21]) AND Data[20]) AND (NOT Data[1])) AND Data[3]) AND Data[2])) OR Data[16])) AND ((NOT ((((Data[21] AND Data[20]) AND (NOT Data[1])) AND Data[3]) AND Data[2])) OR Data[34])) AND ((NOT (((((NOT Data[21]) AND (NOT Data[20])) AND Data[1]) AND Data[3]) AND Data[2])) OR Data[14])) AND ((NOT ((((Data[21] AND (NOT Data[20])) AND Data[1]) AND Data[3]) AND Data[2])) OR Data[17])) AND ((NOT (((((NOT Data[21]) AND Data[20]) AND Data[1]) AND Data[3]) AND Data[2])) OR Data[18])) AND ((NOT ((((Data[21] AND Data[20]) AND Data[1]) AND Data[3]) AND Data[2])) OR Data[19]));
    OutReady := 1;
    CollectInput(RESET:=TRUE);
  END_IF;
END_PROGRAM

CONFIGURATION Config0
  RESOURCE Res0 ON PLC
    TASK task0(INTERVAL := T#20ms,PRIORITY := 0);
    PROGRAM instance0 WITH task0 : Boiler;
  END_RESOURCE
END_CONFIGURATION

(* ---- 5-MUX_heart-pinks-hands.st ---- *)
(*
This code implements a shuffled multiplexer with 5 control bits.
The control bits are: Data[N2], Data[N21], Data[N23], Data[N20], Data[N1]
The input bits are: Data[N5], Data[N25], Data[N4], Data[N3], Data[N27], Data[N22], Data[N24], Data[N26], Data[N31], Data[N8], Data[N29], Data[N30], Data[N35], Data[N6], Data[N7], Data[N9], Data[N10], Data[N15], Data[N32], Data[N28], Data[N11], Data[N36], Data[N12], Data[N14], Data[N13], Data[N16], Data[N34], Data[N33], Data[N37], Data[N18], Data[N17], Data[N19]

The symbolic expression is:
((((((((((((((((((((((((((((((((!(((((!(IN2)) & (!(IN21))) & (!(IN23))) & (!(IN20))) & (!(IN1)))) | IN5) & ((!((((IN2 & (!(IN21))) & (!(IN23))) & (!(IN20))) & (!(IN1)))) | IN25)) & ((!(((((!(IN2)) & IN21) & (!(IN23))) & (!(IN20))) & (!(IN1)))) | IN4)) & ((!((((IN2 & IN21) & (!(IN23))) & (!(IN20))) & (!(IN1)))) | IN3)) & ((!(((((!(IN2)) & (!(IN21))) & IN23) & (!(IN20))) & (!(IN1)))) | IN27)) & ((!((((IN2 & (!(IN21))) & IN23) & (!(IN20))) & (!(IN1)))) | IN22)) & ((!(((((!(IN2)) & IN21) & IN23) & (!(IN20))) & (!(IN1)))) | IN24)) & ((!((((IN2 & IN21) & IN23) & (!(IN20))) & (!(IN1)))) | IN26)) & ((!(((((!(IN2)) & (!(IN21))) & (!(IN23))) & IN20) & (!(IN1)))) | IN31)) & ((!((((IN2 & (!(IN21))) & (!(IN23))) & IN20) & (!(IN1)))) | IN8)) & ((!(((((!(IN2)) & IN21) & (!(IN23))) & IN20) & (!(IN1)))) | IN29)) & ((!((((IN2 & IN21) & (!(IN23))) & IN20) & (!(IN1)))) | IN30)) & ((!(((((!(IN2)) & (!(IN21))) & IN23) & IN20) & (!(IN1)))) | IN35)) & ((!((((IN2 & (!(IN21))) & IN23) & IN20) & (!(IN1)))) | IN6)) & ((!(((((!(IN2)) & IN21) & IN23) & IN20) & (!(IN1)))) | IN7)) & ((!((((IN2 & IN21) & IN23) & IN20) & (!(IN1)))) | IN9)) & ((!(((((!(IN2)) & (!(IN21))) & (!(IN23))) & (!(IN20))) & IN1)) | IN10)) & ((!((((IN2 & (!(IN21))) & (!(IN23))) & (!(IN20))) & IN1)) | IN15)) & ((!(((((!(IN2)) & IN21) & (!(IN23))) & (!(IN20))) & IN1)) | IN32)) & ((!((((IN2 & IN21) & (!(IN23))) & (!(IN20))) & IN1)) | IN28)) & ((!(((((!(IN2)) & (!(IN21))) & IN23) & (!(IN20))) & IN1)) | IN11)) & ((!((((IN2 & (!(IN21))) & IN23) & (!(IN20))) & IN1)) | IN36)) & ((!(((((!(IN2)) & IN21) & IN23) & (!(IN20))) & IN1)) | IN12)) & ((!((((IN2 & IN21) & IN23) & (!(IN20))) & IN1)) | IN14)) & ((!(((((!(IN2)) & (!(IN21))) & (!(IN23))) & IN20) & IN1)) | IN13)) & ((!((((IN2 & (!(IN21))) & (!(IN23))) & IN20) & IN1)) | IN16)) & ((!(((((!(IN2)) & IN21) & (!(IN23))) & IN20) & IN1)) | IN34)) & ((!((((IN2 & IN21) & (!(IN23))) & IN20) & IN1)) | IN33)) & ((!(((((!(IN2)) & (!(IN21))) & IN23) & IN20) & IN1)) | IN37)) & ((!((((IN2 & (!(IN21))) & IN23) & IN20) & IN1)) | IN18)) & ((!(((((!(IN2)) & IN21) & IN23) & IN20) & IN1)) | IN17)) & ((!((((IN2 & IN21) & IN23) & IN20) & IN1)) | IN19)

*)

FUNCTION_BLOCK F_CollectInput
  VAR_IN_OUT
      Data : ARRAY[1..40] OF BOOL;
  END_VAR
  VAR_INPUT
      TICK  : BOOL := 0;
      IN1   : BOOL := 0;
      IN2   : BOOL := 0;
      IN3   : BOOL := 0;
      IN4   : BOOL := 0;
      IN5   : BOOL := 0;
      RESET : BOOL := FALSE;
  END_VAR
  VAR_OUTPUT
      Finished : BOOL;
  END_VAR
  VAR
      j    : USINT := 1;
      tock : BOOL  := 0;
  END_VAR
  IF NOT RESET AND tock = NOT TICK THEN
      Data[j]   := IN1;
      Data[j+1] := IN2;
      Data[j+2] := IN3;
      Data[j+3] := IN4;
      Data[j+4] := IN5;
      j := j + 5;
      tock := TICK;
  ELSE
      j := 1;
      tock := 0;
  END_IF;
  Finished := (j > 40);
END_FUNCTION_BLOCK

PROGRAM Boiler
  VAR
    Data  : ARRAY[1..40] OF BOOL;
    Ready : BOOL;
    CollectInput : F_CollectInput;
  END_VAR
  VAR
    TICK     AT %IX1.0 : BOOL;
    IN1      AT %IX0.3 : BOOL;
    IN2      AT %IX0.4 : BOOL;
    IN3      AT %IX0.5 : BOOL;
    IN4      AT %IX0.6 : BOOL;
    IN5      AT %IX0.7 : BOOL;
    OutReady AT %QX0.0 : BOOL := FALSE;
    FeedNext AT %QX0.1 : BOOL := FALSE;
    Out      AT %QX0.2 : BOOL;
  END_VAR
  CollectInput(TICK:=TICK, IN1:=IN1, IN2:=IN2, IN3:=IN3, IN4:=IN4, IN5:=IN5);
  Ready := CollectInput.Finished;
  FeedNext := 1;
  IF Ready THEN
    Out := (((((((((((((((((((((((((((((((((NOT (((((NOT Data[2]) AND (NOT Data[21])) AND (NOT Data[23])) AND (NOT Data[20])) AND (NOT Data[1]))) OR Data[5]) AND ((NOT ((((Data[2] AND (NOT Data[21])) AND (NOT Data[23])) AND (NOT Data[20])) AND (NOT Data[1]))) OR Data[25])) AND ((NOT (((((NOT Data[2]) AND Data[21]) AND (NOT Data[23])) AND (NOT Data[20])) AND (NOT Data[1]))) OR Data[4])) AND ((NOT ((((Data[2] AND Data[21]) AND (NOT Data[23])) AND (NOT Data[20])) AND (NOT Data[1]))) OR Data[3])) AND ((NOT (((((NOT Data[2]) AND (NOT Data[21])) AND Data[23]) AND (NOT Data[20])) AND (NOT Data[1]))) OR Data[27])) AND ((NOT ((((Data[2] AND (NOT Data[21])) AND Data[23]) AND (NOT Data[20])) AND (NOT Data[1]))) OR Data[22])) AND ((NOT (((((NOT Data[2]) AND Data[21]) AND Data[23]) AND (NOT Data[20])) AND (NOT Data[1]))) OR Data[24])) AND ((NOT ((((Data[2] AND Data[21]) AND Data[23]) AND (NOT Data[20])) AND (NOT Data[1]))) OR Data[26])) AND ((NOT (((((NOT Data[2]) AND (NOT Data[21])) AND (NOT Data[23])) AND Data[20]) AND (NOT Data[1]))) OR Data[31])) AND ((NOT ((((Data[2] AND (NOT Data[21])) AND (NOT Data[23])) AND Data[20]) AND (NOT Data[1]))) OR Data[8])) AND ((NOT (((((NOT Data[2]) AND Data[21]) AND (NOT Data[23])) AND Data[20]) AND (NOT Data[1]))) OR Data[29])) AND ((NOT ((((Data[2] AND Data[21]) AND (NOT Data[23])) AND Data[20]) AND (NOT Data[1]))) OR Data[30])) AND ((NOT (((((NOT Data[2]) AND (NOT Data[21])) AND Data[23]) AND Data[20]) AND (NOT Data[1]))) OR Data[35])) AND ((NOT ((((Data[2] AND (NOT Data[21])) AND Data[23]) AND Data[20]) AND (NOT Data[1]))) OR Data[6])) AND ((NOT (((((NOT Data[2]) AND Data[21]) AND Data[23]) AND Data[20]) AND (NOT Data[1]))) OR Data[7])) AND ((NOT ((((Data[2] AND Data[21]) AND Data[23]) AND Data[20]) AND (NOT Data[1]))) OR Data[9])) AND ((NOT (((((NOT Data[2]) AND (NOT Data[21])) AND (NOT Data[23])) AND (NOT Data[20])) AND Data[1])) OR Data[10])) AND ((NOT ((((Data[2] AND (NOT Data[21])) AND (NOT Data[23])) AND (NOT Data[20])) AND Data[1])) OR Data[15])) AND ((NOT (((((NOT Data[2]) AND Data[21]) AND (NOT Data[23])) AND (NOT Data[20])) AND Data[1])) OR Data[32])) AND ((NOT ((((Data[2] AND Data[21]) AND (NOT Data[23])) AND (NOT Data[20])) AND Data[1])) OR Data[28])) AND ((NOT (((((NOT Data[2]) AND (NOT Data[21])) AND Data[23]) AND (NOT Data[20])) AND Data[1])) OR Data[11])) AND ((NOT ((((Data[2] AND (NOT Data[21])) AND Data[23]) AND (NOT Data[20])) AND Data[1])) OR Data[36])) AND ((NOT (((((NOT Data[2]) AND Data[21]) AND Data[23]) AND (NOT Data[20])) AND Data[1])) OR Data[12])) AND ((NOT ((((Data[2] AND Data[21]) AND Data[23]) AND (NOT Data[20])) AND Data[1])) OR Data[14])) AND ((NOT (((((NOT Data[2]) AND (NOT Data[21])) AND (NOT Data[23])) AND Data[20]) AND Data[1])) OR Data[13])) AND ((NOT ((((Data[2] AND (NOT Data[21])) AND (NOT Data[23])) AND Data[20]) AND Data[1])) OR Data[16])) AND ((NOT (((((NOT Data[2]) AND Data[21]) AND (NOT Data[23])) AND Data[20]) AND Data[1])) OR Data[34])) AND ((NOT ((((Data[2] AND Data[21]) AND (NOT Data[23])) AND Data[20]) AND Data[1])) OR Data[33])) AND ((NOT (((((NOT Data[2]) AND (NOT Data[21])) AND Data[23]) AND Data[20]) AND Data[1])) OR Data[37])) AND ((NOT ((((Data[2] AND (NOT Data[21])) AND Data[23]) AND Data[20]) AND Data[1])) OR Data[18])) AND ((NOT (((((NOT Data[2]) AND Data[21]) AND Data[23]) AND Data[20]) AND Data[1])) OR Data[17])) AND ((NOT ((((Data[2] AND Data[21]) AND Data[23]) AND Data[20]) AND Data[1])) OR Data[19]));
    OutReady := 1;
    CollectInput(RESET:=TRUE);
  END_IF;
END_PROGRAM

CONFIGURATION Config0
  RESOURCE Res0 ON PLC
    TASK task0(INTERVAL := T#20ms,PRIORITY := 0);
    PROGRAM instance0 WITH task0 : Boiler;
  END_RESOURCE
END_CONFIGURATION

(* ---- 5-MUX_homos-bakes-madam.st ---- *)
(*
This code implements a shuffled multiplexer with 5 control bits.
The control bits are: Data[N2], Data[N21], Data[N24], Data[N20], Data[N25]
The input bits are: Data[N26], Data[N22], Data[N27], Data[N28], Data[N31], Data[N23], Data[N3], Data[N1], Data[N30], Data[N4], Data[N29], Data[N32], Data[N5], Data[N34], Data[N33], Data[N35], Data[N6], Data[N36], Data[N37], Data[N7], Data[N12], Data[N8], Data[N9], Data[N10], Data[N11], Data[N13], Data[N14], Data[N15], Data[N19], Data[N16], Data[N17], Data[N18]

The symbolic expression is:
((((((((((((((((((((((((((((((((!(((((!(IN2)) & (!(IN21))) & (!(IN24))) & (!(IN20))) & (!(IN25)))) | IN26) & ((!((((IN2 & (!(IN21))) & (!(IN24))) & (!(IN20))) & (!(IN25)))) | IN22)) & ((!(((((!(IN2)) & IN21) & (!(IN24))) & (!(IN20))) & (!(IN25)))) | IN27)) & ((!((((IN2 & IN21) & (!(IN24))) & (!(IN20))) & (!(IN25)))) | IN28)) & ((!(((((!(IN2)) & (!(IN21))) & IN24) & (!(IN20))) & (!(IN25)))) | IN31)) & ((!((((IN2 & (!(IN21))) & IN24) & (!(IN20))) & (!(IN25)))) | IN23)) & ((!(((((!(IN2)) & IN21) & IN24) & (!(IN20))) & (!(IN25)))) | IN3)) & ((!((((IN2 & IN21) & IN24) & (!(IN20))) & (!(IN25)))) | IN1)) & ((!(((((!(IN2)) & (!(IN21))) & (!(IN24))) & IN20) & (!(IN25)))) | IN30)) & ((!((((IN2 & (!(IN21))) & (!(IN24))) & IN20) & (!(IN25)))) | IN4)) & ((!(((((!(IN2)) & IN21) & (!(IN24))) & IN20) & (!(IN25)))) | IN29)) & ((!((((IN2 & IN21) & (!(IN24))) & IN20) & (!(IN25)))) | IN32)) & ((!(((((!(IN2)) & (!(IN21))) & IN24) & IN20) & (!(IN25)))) | IN5)) & ((!((((IN2 & (!(IN21))) & IN24) & IN20) & (!(IN25)))) | IN34)) & ((!(((((!(IN2)) & IN21) & IN24) & IN20) & (!(IN25)))) | IN33)) & ((!((((IN2 & IN21) & IN24) & IN20) & (!(IN25)))) | IN35)) & ((!(((((!(IN2)) & (!(IN21))) & (!(IN24))) & (!(IN20))) & IN25)) | IN6)) & ((!((((IN2 & (!(IN21))) & (!(IN24))) & (!(IN20))) & IN25)) | IN36)) & ((!(((((!(IN2)) & IN21) & (!(IN24))) & (!(IN20))) & IN25)) | IN37)) & ((!((((IN2 & IN21) & (!(IN24))) & (!(IN20))) & IN25)) | IN7)) & ((!(((((!(IN2)) & (!(IN21))) & IN24) & (!(IN20))) & IN25)) | IN12)) & ((!((((IN2 & (!(IN21))) & IN24) & (!(IN20))) & IN25)) | IN8)) & ((!(((((!(IN2)) & IN21) & IN24) & (!(IN20))) & IN25)) | IN9)) & ((!((((IN2 & IN21) & IN24) & (!(IN20))) & IN25)) | IN10)) & ((!(((((!(IN2)) & (!(IN21))) & (!(IN24))) & IN20) & IN25)) | IN11)) & ((!((((IN2 & (!(IN21))) & (!(IN24))) & IN20) & IN25)) | IN13)) & ((!(((((!(IN2)) & IN21) & (!(IN24))) & IN20) & IN25)) | IN14)) & ((!((((IN2 & IN21) & (!(IN24))) & IN20) & IN25)) | IN15)) & ((!(((((!(IN2)) & (!(IN21))) & IN24) & IN20) & IN25)) | IN19)) & ((!((((IN2 & (!(IN21))) & IN24) & IN20) & IN25)) | IN16)) & ((!(((((!(IN2)) & IN21) & IN24) & IN20) & IN25)) | IN17)) & ((!((((IN2 & IN21) & IN24) & IN20) & IN25)) | IN18)

*)

FUNCTION_BLOCK F_CollectInput
  VAR_IN_OUT
      Data : ARRAY[1..40] OF BOOL;
  END_VAR
  VAR_INPUT
      TICK  : BOOL := 0;
      IN1   : BOOL := 0;
      IN2   : BOOL := 0;
      IN3   : BOOL := 0;
      IN4   : BOOL := 0;
      IN5   : BOOL := 0;
      RESET : BOOL := FALSE;
  END_VAR
  VAR_OUTPUT
      Finished : BOOL;
  END_VAR
  VAR
      j    : USINT := 1;
      tock : BOOL  := 0;
  END_VAR
  IF NOT RESET AND tock = NOT TICK THEN
      Data[j]   := IN1;
      Data[j+1] := IN2;
      Data[j+2] := IN3;
      Data[j+3] := IN4;
      Data[j+4] := IN5;
      j := j + 5;
      tock := TICK;
  ELSE
      j := 1;
      tock := 0;
  END_IF;
  Finished := (j > 40);
END_FUNCTION_BLOCK

PROGRAM Boiler
  VAR
    Data  : ARRAY[1..40] OF BOOL;
    Ready : BOOL;
    CollectInput : F_CollectInput;
  END_VAR
  VAR
    TICK     AT %IX1.0 : BOOL;
    IN1      AT %IX0.3 : BOOL;
    IN2      AT %IX0.4 : BOOL;
    IN3      AT %IX0.5 : BOOL;
    IN4      AT %IX0.6 : BOOL;
    IN5      AT %IX0.7 : BOOL;
    OutReady AT %QX0.0 : BOOL := FALSE;
    FeedNext AT %QX0.1 : BOOL := FALSE;
    Out      AT %QX0.2 : BOOL;
  END_VAR
  CollectInput(TICK:=TICK, IN1:=IN1, IN2:=IN2, IN3:=IN3, IN4:=IN4, IN5:=IN5);
  Ready := CollectInput.Finished;
  FeedNext := 1;
  IF Ready THEN
    Out := (((((((((((((((((((((((((((((((((NOT (((((NOT Data[2]) AND (NOT Data[21])) AND (NOT Data[24])) AND (NOT Data[20])) AND (NOT Data[25]))) OR Data[26]) AND ((NOT ((((Data[2] AND (NOT Data[21])) AND (NOT Data[24])) AND (NOT Data[20])) AND (NOT Data[25]))) OR Data[22])) AND ((NOT (((((NOT Data[2]) AND Data[21]) AND (NOT Data[24])) AND (NOT Data[20])) AND (NOT Data[25]))) OR Data[27])) AND ((NOT ((((Data[2] AND Data[21]) AND (NOT Data[24])) AND (NOT Data[20])) AND (NOT Data[25]))) OR Data[28])) AND ((NOT (((((NOT Data[2]) AND (NOT Data[21])) AND Data[24]) AND (NOT Data[20])) AND (NOT Data[25]))) OR Data[31])) AND ((NOT ((((Data[2] AND (NOT Data[21])) AND Data[24]) AND (NOT Data[20])) AND (NOT Data[25]))) OR Data[23])) AND ((NOT (((((NOT Data[2]) AND Data[21]) AND Data[24]) AND (NOT Data[20])) AND (NOT Data[25]))) OR Data[3])) AND ((NOT ((((Data[2] AND Data[21]) AND Data[24]) AND (NOT Data[20])) AND (NOT Data[25]))) OR Data[1])) AND ((NOT (((((NOT Data[2]) AND (NOT Data[21])) AND (NOT Data[24])) AND Data[20]) AND (NOT Data[25]))) OR Data[30])) AND ((NOT ((((Data[2] AND (NOT Data[21])) AND (NOT Data[24])) AND Data[20]) AND (NOT Data[25]))) OR Data[4])) AND ((NOT (((((NOT Data[2]) AND Data[21]) AND (NOT Data[24])) AND Data[20]) AND (NOT Data[25]))) OR Data[29])) AND ((NOT ((((Data[2] AND Data[21]) AND (NOT Data[24])) AND Data[20]) AND (NOT Data[25]))) OR Data[32])) AND ((NOT (((((NOT Data[2]) AND (NOT Data[21])) AND Data[24]) AND Data[20]) AND (NOT Data[25]))) OR Data[5])) AND ((NOT ((((Data[2] AND (NOT Data[21])) AND Data[24]) AND Data[20]) AND (NOT Data[25]))) OR Data[34])) AND ((NOT (((((NOT Data[2]) AND Data[21]) AND Data[24]) AND Data[20]) AND (NOT Data[25]))) OR Data[33])) AND ((NOT ((((Data[2] AND Data[21]) AND Data[24]) AND Data[20]) AND (NOT Data[25]))) OR Data[35])) AND ((NOT (((((NOT Data[2]) AND (NOT Data[21])) AND (NOT Data[24])) AND (NOT Data[20])) AND Data[25])) OR Data[6])) AND ((NOT ((((Data[2] AND (NOT Data[21])) AND (NOT Data[24])) AND (NOT Data[20])) AND Data[25])) OR Data[36])) AND ((NOT (((((NOT Data[2]) AND Data[21]) AND (NOT Data[24])) AND (NOT Data[20])) AND Data[25])) OR Data[37])) AND ((NOT ((((Data[2] AND Data[21]) AND (NOT Data[24])) AND (NOT Data[20])) AND Data[25])) OR Data[7])) AND ((NOT (((((NOT Data[2]) AND (NOT Data[21])) AND Data[24]) AND (NOT Data[20])) AND Data[25])) OR Data[12])) AND ((NOT ((((Data[2] AND (NOT Data[21])) AND Data[24]) AND (NOT Data[20])) AND Data[25])) OR Data[8])) AND ((NOT (((((NOT Data[2]) AND Data[21]) AND Data[24]) AND (NOT Data[20])) AND Data[25])) OR Data[9])) AND ((NOT ((((Data[2] AND Data[21]) AND Data[24]) AND (NOT Data[20])) AND Data[25])) OR Data[10])) AND ((NOT (((((NOT Data[2]) AND (NOT Data[21])) AND (NOT Data[24])) AND Data[20]) AND Data[25])) OR Data[11])) AND ((NOT ((((Data[2] AND (NOT Data[21])) AND (NOT Data[24])) AND Data[20]) AND Data[25])) OR Data[13])) AND ((NOT (((((NOT Data[2]) AND Data[21]) AND (NOT Data[24])) AND Data[20]) AND Data[25])) OR Data[14])) AND ((NOT ((((Data[2] AND Data[21]) AND (NOT Data[24])) AND Data[20]) AND Data[25])) OR Data[15])) AND ((NOT (((((NOT Data[2]) AND (NOT Data[21])) AND Data[24]) AND Data[20]) AND Data[25])) OR Data[19])) AND ((NOT ((((Data[2] AND (NOT Data[21])) AND Data[24]) AND Data[20]) AND Data[25])) OR Data[16])) AND ((NOT (((((NOT Data[2]) AND Data[21]) AND Data[24]) AND Data[20]) AND Data[25])) OR Data[17])) AND ((NOT ((((Data[2] AND Data[21]) AND Data[24]) AND Data[20]) AND Data[25])) OR Data[18]));
    OutReady := 1;
    CollectInput(RESET:=TRUE);
  END_IF;
END_PROGRAM

CONFIGURATION Config0
  RESOURCE Res0 ON PLC
    TASK task0(INTERVAL := T#20ms,PRIORITY := 0);
    PROGRAM instance0 WITH task0 : Boiler;
  END_RESOURCE
END_CONFIGURATION

(* ---- 5-MUX_horse-peers-edges.st ---- *)
(*
This code implements a shuffled multiplexer with 5 control bits.
The control bits are: Data[N20], Data[N22], Data[N21], Data[N3], Data[N1]
The input bits are: Data[N5], Data[N2], Data[N24], Data[N6], Data[N4], Data[N23], Data[N7], Data[N27], Data[N10], Data[N8], Data[N25], Data[N26], Data[N29], Data[N9], Data[N12], Data[N28], Data[N33], Data[N30], Data[N31], Data[N36], Data[N11], Data[N32], Data[N34], Data[N13], Data[N15], Data[N37], Data[N35], Data[N16], Data[N17], Data[N14], Data[N18], Data[N19]

The symbolic expression is:
((((((((((((((((((((((((((((((((!(((((!(IN20)) & (!(IN22))) & (!(IN21))) & (!(IN3))) & (!(IN1)))) | IN5) & ((!((((IN20 & (!(IN22))) & (!(IN21))) & (!(IN3))) & (!(IN1)))) | IN2)) & ((!(((((!(IN20)) & IN22) & (!(IN21))) & (!(IN3))) & (!(IN1)))) | IN24)) & ((!((((IN20 & IN22) & (!(IN21))) & (!(IN3))) & (!(IN1)))) | IN6)) & ((!(((((!(IN20)) & (!(IN22))) & IN21) & (!(IN3))) & (!(IN1)))) | IN4)) & ((!((((IN20 & (!(IN22))) & IN21) & (!(IN3))) & (!(IN1)))) | IN23)) & ((!(((((!(IN20)) & IN22) & IN21) & (!(IN3))) & (!(IN1)))) | IN7)) & ((!((((IN20 & IN22) & IN21) & (!(IN3))) & (!(IN1)))) | IN27)) & ((!(((((!(IN20)) & (!(IN22))) & (!(IN21))) & IN3) & (!(IN1)))) | IN10)) & ((!((((IN20 & (!(IN22))) & (!(IN21))) & IN3) & (!(IN1)))) | IN8)) & ((!(((((!(IN20)) & IN22) & (!(IN21))) & IN3) & (!(IN1)))) | IN25)) & ((!((((IN20 & IN22) & (!(IN21))) & IN3) & (!(IN1)))) | IN26)) & ((!(((((!(IN20)) & (!(IN22))) & IN21) & IN3) & (!(IN1)))) | IN29)) & ((!((((IN20 & (!(IN22))) & IN21) & IN3) & (!(IN1)))) | IN9)) & ((!(((((!(IN20)) & IN22) & IN21) & IN3) & (!(IN1)))) | IN12)) & ((!((((IN20 & IN22) & IN21) & IN3) & (!(IN1)))) | IN28)) & ((!(((((!(IN20)) & (!(IN22))) & (!(IN21))) & (!(IN3))) & IN1)) | IN33)) & ((!((((IN20 & (!(IN22))) & (!(IN21))) & (!(IN3))) & IN1)) | IN30)) & ((!(((((!(IN20)) & IN22) & (!(IN21))) & (!(IN3))) & IN1)) | IN31)) & ((!((((IN20 & IN22) & (!(IN21))) & (!(IN3))) & IN1)) | IN36)) & ((!(((((!(IN20)) & (!(IN22))) & IN21) & (!(IN3))) & IN1)) | IN11)) & ((!((((IN20 & (!(IN22))) & IN21) & (!(IN3))) & IN1)) | IN32)) & ((!(((((!(IN20)) & IN22) & IN21) & (!(IN3))) & IN1)) | IN34)) & ((!((((IN20 & IN22) & IN21) & (!(IN3))) & IN1)) | IN13)) & ((!(((((!(IN20)) & (!(IN22))) & (!(IN21))) & IN3) & IN1)) | IN15)) & ((!((((IN20 & (!(IN22))) & (!(IN21))) & IN3) & IN1)) | IN37)) & ((!(((((!(IN20)) & IN22) & (!(IN21))) & IN3) & IN1)) | IN35)) & ((!((((IN20 & IN22) & (!(IN21))) & IN3) & IN1)) | IN16)) & ((!(((((!(IN20)) & (!(IN22))) & IN21) & IN3) & IN1)) | IN17)) & ((!((((IN20 & (!(IN22))) & IN21) & IN3) & IN1)) | IN14)) & ((!(((((!(IN20)) & IN22) & IN21) & IN3) & IN1)) | IN18)) & ((!((((IN20 & IN22) & IN21) & IN3) & IN1)) | IN19)

*)

FUNCTION_BLOCK F_CollectInput
  VAR_IN_OUT
      Data : ARRAY[1..40] OF BOOL;
  END_VAR
  VAR_INPUT
      TICK  : BOOL := 0;
      IN1   : BOOL := 0;
      IN2   : BOOL := 0;
      IN3   : BOOL := 0;
      IN4   : BOOL := 0;
      IN5   : BOOL := 0;
      RESET : BOOL := FALSE;
  END_VAR
  VAR_OUTPUT
      Finished : BOOL;
  END_VAR
  VAR
      j    : USINT := 1;
      tock : BOOL  := 0;
  END_VAR
  IF NOT RESET AND tock = NOT TICK THEN
      Data[j]   := IN1;
      Data[j+1] := IN2;
      Data[j+2] := IN3;
      Data[j+3] := IN4;
      Data[j+4] := IN5;
      j := j + 5;
      tock := TICK;
  ELSE
      j := 1;
      tock := 0;
  END_IF;
  Finished := (j > 40);
END_FUNCTION_BLOCK

PROGRAM Boiler
  VAR
    Data  : ARRAY[1..40] OF BOOL;
    Ready : BOOL;
    CollectInput : F_CollectInput;
  END_VAR
  VAR
    TICK     AT %IX1.0 : BOOL;
    IN1      AT %IX0.3 : BOOL;
    IN2      AT %IX0.4 : BOOL;
    IN3      AT %IX0.5 : BOOL;
    IN4      AT %IX0.6 : BOOL;
    IN5      AT %IX0.7 : BOOL;
    OutReady AT %QX0.0 : BOOL := FALSE;
    FeedNext AT %QX0.1 : BOOL := FALSE;
    Out      AT %QX0.2 : BOOL;
  END_VAR
  CollectInput(TICK:=TICK, IN1:=IN1, IN2:=IN2, IN3:=IN3, IN4:=IN4, IN5:=IN5);
  Ready := CollectInput.Finished;
  FeedNext := 1;
  IF Ready THEN
    Out := (((((((((((((((((((((((((((((((((NOT (((((NOT Data[20]) AND (NOT Data[22])) AND (NOT Data[21])) AND (NOT Data[3])) AND (NOT Data[1]))) OR Data[5]) AND ((NOT ((((Data[20] AND (NOT Data[22])) AND (NOT Data[21])) AND (NOT Data[3])) AND (NOT Data[1]))) OR Data[2])) AND ((NOT (((((NOT Data[20]) AND Data[22]) AND (NOT Data[21])) AND (NOT Data[3])) AND (NOT Data[1]))) OR Data[24])) AND ((NOT ((((Data[20] AND Data[22]) AND (NOT Data[21])) AND (NOT Data[3])) AND (NOT Data[1]))) OR Data[6])) AND ((NOT (((((NOT Data[20]) AND (NOT Data[22])) AND Data[21]) AND (NOT Data[3])) AND (NOT Data[1]))) OR Data[4])) AND ((NOT ((((Data[20] AND (NOT Data[22])) AND Data[21]) AND (NOT Data[3])) AND (NOT Data[1]))) OR Data[23])) AND ((NOT (((((NOT Data[20]) AND Data[22]) AND Data[21]) AND (NOT Data[3])) AND (NOT Data[1]))) OR Data[7])) AND ((NOT ((((Data[20] AND Data[22]) AND Data[21]) AND (NOT Data[3])) AND (NOT Data[1]))) OR Data[27])) AND ((NOT (((((NOT Data[20]) AND (NOT Data[22])) AND (NOT Data[21])) AND Data[3]) AND (NOT Data[1]))) OR Data[10])) AND ((NOT ((((Data[20] AND (NOT Data[22])) AND (NOT Data[21])) AND Data[3]) AND (NOT Data[1]))) OR Data[8])) AND ((NOT (((((NOT Data[20]) AND Data[22]) AND (NOT Data[21])) AND Data[3]) AND (NOT Data[1]))) OR Data[25])) AND ((NOT ((((Data[20] AND Data[22]) AND (NOT Data[21])) AND Data[3]) AND (NOT Data[1]))) OR Data[26])) AND ((NOT (((((NOT Data[20]) AND (NOT Data[22])) AND Data[21]) AND Data[3]) AND (NOT Data[1]))) OR Data[29])) AND ((NOT ((((Data[20] AND (NOT Data[22])) AND Data[21]) AND Data[3]) AND (NOT Data[1]))) OR Data[9])) AND ((NOT (((((NOT Data[20]) AND Data[22]) AND Data[21]) AND Data[3]) AND (NOT Data[1]))) OR Data[12])) AND ((NOT ((((Data[20] AND Data[22]) AND Data[21]) AND Data[3]) AND (NOT Data[1]))) OR Data[28])) AND ((NOT (((((NOT Data[20]) AND (NOT Data[22])) AND (NOT Data[21])) AND (NOT Data[3])) AND Data[1])) OR Data[33])) AND ((NOT ((((Data[20] AND (NOT Data[22])) AND (NOT Data[21])) AND (NOT Data[3])) AND Data[1])) OR Data[30])) AND ((NOT (((((NOT Data[20]) AND Data[22]) AND (NOT Data[21])) AND (NOT Data[3])) AND Data[1])) OR Data[31])) AND ((NOT ((((Data[20] AND Data[22]) AND (NOT Data[21])) AND (NOT Data[3])) AND Data[1])) OR Data[36])) AND ((NOT (((((NOT Data[20]) AND (NOT Data[22])) AND Data[21]) AND (NOT Data[3])) AND Data[1])) OR Data[11])) AND ((NOT ((((Data[20] AND (NOT Data[22])) AND Data[21]) AND (NOT Data[3])) AND Data[1])) OR Data[32])) AND ((NOT (((((NOT Data[20]) AND Data[22]) AND Data[21]) AND (NOT Data[3])) AND Data[1])) OR Data[34])) AND ((NOT ((((Data[20] AND Data[22]) AND Data[21]) AND (NOT Data[3])) AND Data[1])) OR Data[13])) AND ((NOT (((((NOT Data[20]) AND (NOT Data[22])) AND (NOT Data[21])) AND Data[3]) AND Data[1])) OR Data[15])) AND ((NOT ((((Data[20] AND (NOT Data[22])) AND (NOT Data[21])) AND Data[3]) AND Data[1])) OR Data[37])) AND ((NOT (((((NOT Data[20]) AND Data[22]) AND (NOT Data[21])) AND Data[3]) AND Data[1])) OR Data[35])) AND ((NOT ((((Data[20] AND Data[22]) AND (NOT Data[21])) AND Data[3]) AND Data[1])) OR Data[16])) AND ((NOT (((((NOT Data[20]) AND (NOT Data[22])) AND Data[21]) AND Data[3]) AND Data[1])) OR Data[17])) AND ((NOT ((((Data[20] AND (NOT Data[22])) AND Data[21]) AND Data[3]) AND Data[1])) OR Data[14])) AND ((NOT (((((NOT Data[20]) AND Data[22]) AND Data[21]) AND Data[3]) AND Data[1])) OR Data[18])) AND ((NOT ((((Data[20] AND Data[22]) AND Data[21]) AND Data[3]) AND Data[1])) OR Data[19]));
    OutReady := 1;
    CollectInput(RESET:=TRUE);
  END_IF;
END_PROGRAM

CONFIGURATION Config0
  RESOURCE Res0 ON PLC
    TASK task0(INTERVAL := T#20ms,PRIORITY := 0);
    PROGRAM instance0 WITH task0 : Boiler;
  END_RESOURCE
END_CONFIGURATION
